    RC2_Transmit_PDO_Mapping_StatusWord_6041_00 : UINT;
    RC2_Transmit_PDO_Mapping_Position_actual_value_6064_00 : DINT;
    RC2_Transmit_PDO_Mapping_Mode_of_operation_display_6061_00 : SINT;
    RC2_Transmit_PDO_Mapping_Following_error_actual_valu_60F4_00 : DINT;
    RC2_Transmit_PDO_Mapping_Torque_actual_value_6077_00 : INT;
    RC2_Transmit_PDO_Mapping_Digital_inputs_60FD_00 : UDINT;
    RC2_Transmit_PDO_Mapping_Error_code_603F_00 : UINT;
    RC3_Receive_PDO_Mapping_ControlWord_6040_00 : UINT;
    RC3_Receive_PDO_Mapping_Target_Position_607A_00 : DINT;
    RC3_Receive_PDO_Mapping_Mode_of_operation_6060_00 : SINT;
    RC3_Receive_PDO_Mapping_Profile_velocity_6081_00 : UDINT;
    RC3_Receive_PDO_Mapping_Profile_acceleration_6083_00 : UDINT;
    RC3_Receive_PDO_Mapping_Profile_deceleration_6084_00 : UDINT;
    RC3_Receive_PDO_Mapping_Physical_outputs_60FE_01 : UDINT;
    RC3_Transmit_PDO_Mapping_StatusWord_6041_00 : UINT;
    RC3_Transmit_PDO_Mapping_Position_actual_value_6064_00 : DINT;
    RC3_Transmit_PDO_Mapping_Mode_of_operation_display_6061_00 : SINT;
    RC3_Transmit_PDO_Mapping_Following_error_actual_valu_60F4_00 : DINT;
    RC3_Transmit_PDO_Mapping_Torque_actual_value_6077_00 : INT;
    RC3_Transmit_PDO_Mapping_Digital_inputs_60FD_00 : UDINT;
    RC3_Transmit_PDO_Mapping_Error_code_603F_00 : UINT;
    RC4_Receive_PDO_Mapping_ControlWord_6040_00 : UINT;
    RC4_Receive_PDO_Mapping_Target_Position_607A_00 : DINT;
    RC4_Receive_PDO_Mapping_Mode_of_operation_6060_00 : SINT;
    RC4_Receive_PDO_Mapping_Profile_velocity_6081_00 : UDINT;
    RC4_Receive_PDO_Mapping_Profile_acceleration_6083_00 : UDINT;
    RC4_Receive_PDO_Mapping_Profile_deceleration_6084_00 : UDINT;
    RC4_Receive_PDO_Mapping_Physical_outputs_60FE_01 : UDINT;
    RC4_Transmit_PDO_Mapping_StatusWord_6041_00 : UINT;
    RC4_Transmit_PDO_Mapping_Position_actual_value_6064_00 : DINT;
    RC4_Transmit_PDO_Mapping_Mode_of_operation_display_6061_00 : SINT;
    RC4_Transmit_PDO_Mapping_Following_error_actual_valu_60F4_00 : DINT;
    RC4_Transmit_PDO_Mapping_Torque_actual_value_6077_00 : INT;
    RC4_Transmit_PDO_Mapping_Digital_inputs_60FD_00 : UDINT;
    RC4_Transmit_PDO_Mapping_Error_code_603F_00 : UINT;
    RC5_Receive_PDO_Mapping_ControlWord_6040_00 : UINT;
    RC5_Receive_PDO_Mapping_Target_Position_607A_00 : DINT;
    RC5_Receive_PDO_Mapping_Mode_of_operation_6060_00 : SINT;
    RC5_Receive_PDO_Mapping_Profile_velocity_6081_00 : UDINT;
    RC5_Receive_PDO_Mapping_Profile_acceleration_6083_00 : UDINT;
    RC5_Receive_PDO_Mapping_Profile_deceleration_6084_00 : UDINT;
    RC5_Receive_PDO_Mapping_Physical_outputs_60FE_01 : UDINT;
    RC5_Transmit_PDO_Mapping_StatusWord_6041_00 : UINT;
    RC5_Transmit_PDO_Mapping_Position_actual_value_6064_00 : DINT;
    RC5_Transmit_PDO_Mapping_Mode_of_operation_display_6061_00 : SINT;
    RC5_Transmit_PDO_Mapping_Following_error_actual_valu_60F4_00 : DINT;
    RC5_Transmit_PDO_Mapping_Torque_actual_value_6077_00 : INT;
    RC5_Transmit_PDO_Mapping_Digital_inputs_60FD_00 : UDINT;
    RC5_Transmit_PDO_Mapping_Error_code_603F_00 : UINT;
    RC6_Receive_PDO_Mapping_ControlWord_6040_00 : UINT;
    RC6_Receive_PDO_Mapping_ControlWord_6040_00_1 : UINT;
    RC6_Receive_PDO_Mapping_Target_Position_607A_00 : DINT;
    RC6_Receive_PDO_Mapping_Mode_of_operation_6060_00 : SINT;
    RC6_Receive_PDO_Mapping_Profile_velocity_6081_00 : UDINT;
    RC6_Receive_PDO_Mapping_Profile_acceleration_6083_00 : UDINT;
    RC6_Receive_PDO_Mapping_Profile_deceleration_6084_00 : UDINT;
    RC6_Receive_PDO_Mapping_Physical_outputs_60FE_01 : UDINT;
    RC6_Transmit_PDO_Mapping_StatusWord_6041_00 : UINT;
    RC6_Transmit_PDO_Mapping_Position_actual_value_6064_00 : DINT;
    RC6_Transmit_PDO_Mapping_Mode_of_operation_display_6061_00 : SINT;
    RC6_Transmit_PDO_Mapping_Following_error_actual_valu_60F4_00 : DINT;
    RC6_Transmit_PDO_Mapping_Torque_actual_value_6077_00 : INT;
    RC6_Transmit_PDO_Mapping_Digital_inputs_60FD_00 : UDINT;
    RC6_Transmit_PDO_Mapping_Error_code_603F_00 : UINT;
END_VAR
VAR_GLOBAL RETAIN
    RCON1_OUT : ARRAY[1..6] OF ST_RCON_Direct_OUT_Axis;  (* #RCON1 出力値; [2] #B(右側) NG1排出(上下); [3] #A(左側) SF/NG2仕分け(左右); [4] #B(右側) SF/NG2排出(送り); [5] #A(左側) SF/NG2排出(上下); [6] #B(右側) SF/NG2排出(上下); [1].Control.Pause 一時停止（安全停止とは別）（未接続）; [1] #A(左側) NG1排出(上下); [1].TargetPos_mm 目標位置 [mm]; [1].PositionBand_mm 位置決め幅 [mm]; [1].Speed_mm_s 指令速度 [mm/s]; [1].AccDec_G 加減速度 [G]; [1].PushLimit_pct 押付け制限 [%]（未使用）; [1].Control.Start 移動開始; [1].Control.Home 原点復帰（未接続）; [1].Control.Reset 異常リセット; [1].Control.ServoOn サーボON; [1].Control.InchingSelect インチング選択（OFF=ジョグ）; [1].Control.JogSpeedSelect ジョグ速度切替（未接続）; [1].Control.JogMinus 原点方向ジョグ（未接続）; [1].Control.JogPlus 反原点方向ジョグ（未接続）; [1].Control.GainSelect0 ゲイン選択0（未使用）; [1].Control.GainSelect1 ゲイン選択1（未使用）; [1].Control.PushEnable 押付け選択（OFF=位置決め）（未使用）; [1].Control.PushDirection 押付け方向（未使用）; [1].Control.RelativeMove 相対移動（OFF=絶対）（未使用）; [1].Control.BrakeRelease ブレーキ強制解除（落下注意）; [2].TargetPos_mm 目標位置 [mm]; [2].PositionBand_mm 位置決め幅 [mm]; [2].Speed_mm_s 指令速度 [mm/s]; [2].AccDec_G 加減速度 [G]; [2].PushLimit_pct 押付け制限 [%]（未使用）; [2].Control.Start 移動開始; [2].Control.Home 原点復帰（未接続）; [2].Control.Pause 一時停止（安全停止とは別）（未接続）; [2].Control.Reset 異常リセット; [2].Control.ServoOn サーボON; [2].Control.InchingSelect インチング選択（OFF=ジョグ）; [2].Control.JogSpeedSelect ジョグ速度切替（未接続）; [2].Control.JogMinus 原点方向ジョグ（未接続）; [2].Control.JogPlus 反原点方向ジョグ（未接続）; [2].Control.GainSelect0 ゲイン選択0（未使用）; [2].Control.GainSelect1 ゲイン選択1（未使用）; [2].Control.PushEnable 押付け選択（OFF=位置決め）（未使用）; [2].Control.PushDirection 押付け方向（未使用）; [2].Control.RelativeMove 相対移動（OFF=絶対）（未使用）; [2].Control.BrakeRelease ブレーキ強制解除（落下注意）; [3].TargetPos_mm 目標位置 [mm]; [3].PositionBand_mm 位置決め幅 [mm]; [3].Speed_mm_s 指令速度 [mm/s]; [3].AccDec_G 加減速度 [G]; [3].PushLimit_pct 押付け制限 [%]（未使用）; [3].Control.Start 移動開始; [3].Control.Home 原点復帰（未接続）; [3].Control.Pause 一時停止（安全停止とは別）（未接続）; [3].Control.Reset 異常リセット; [3].Control.ServoOn サーボON; [3].Control.InchingSelect インチング選択（OFF=ジョグ）; [3].Control.JogSpeedSelect ジョグ速度切替（未接続）; [3].Control.JogMinus 原点方向ジョグ（未接続）; [3].Control.JogPlus 反原点方向ジョグ（未接続）; [3].Control.GainSelect0 ゲイン選択0（未使用）; [3].Control.GainSelect1 ゲイン選択1（未使用）; [3].Control.PushEnable 押付け選択（OFF=位置決め）（未使用）; [3].Control.PushDirection 押付け方向（未使用）; [3].Control.RelativeMove 相対移動（OFF=絶対）（未使用）; [3].Control.BrakeRelease ブレーキ強制解除（落下注意）; [4].TargetPos_mm 目標位置 [mm]; [4].PositionBand_mm 位置決め幅 [mm]; [4].Speed_mm_s 指令速度 [mm/s]; [4].AccDec_G 加減速度 [G]; [4].PushLimit_pct 押付け制限 [%]（未使用）; [4].Control.Start 移動開始; [4].Control.Home 原点復帰（未接続）; [4].Control.Pause 一時停止（安全停止とは別）（未接続）; [4].Control.Reset 異常リセット; [4].Control.ServoOn サーボON; [4].Control.InchingSelect インチング選択（OFF=ジョグ）; [4].Control.JogSpeedSelect ジョグ速度切替（未接続）; [4].Control.JogMinus 原点方向ジョグ（未接続）; [4].Control.JogPlus 反原点方向ジョグ（未接続）; [4].Control.GainSelect0 ゲイン選択0（未使用）; [4].Control.GainSelect1 ゲイン選択1（未使用）; [4].Control.PushEnable 押付け選択（OFF=位置決め）（未使用）; [4].Control.PushDirection 押付け方向（未使用）; [4].Control.RelativeMove 相対移動（OFF=絶対）（未使用）; [4].Control.BrakeRelease ブレーキ強制解除（落下注意）; [5].TargetPos_mm 目標位置 [mm]; [5].PositionBand_mm 位置決め幅 [mm]; [5].Speed_mm_s 指令速度 [mm/s]; [5].AccDec_G 加減速度 [G]; [5].PushLimit_pct 押付け制限 [%]（未使用）; [5].Control.Start 移動開始; [5].Control.Home 原点復帰（未接続）; [5].Control.Pause 一時停止（安全停止とは別）（未接続）; [5].Control.Reset 異常リセット; [5].Control.ServoOn サーボON; [5].Control.InchingSelect インチング選択（OFF=ジョグ）; [5].Control.JogSpeedSelect ジョグ速度切替（未接続）; [5].Control.JogMinus 原点方向ジョグ（未接続）; [5].Control.JogPlus 反原点方向ジョグ（未接続）; [5].Control.GainSelect0 ゲイン選択0（未使用）; [5].Control.GainSelect1 ゲイン選択1（未使用）; [5].Control.PushEnable 押付け選択（OFF=位置決め）（未使用）; [5].Control.PushDirection 押付け方向（未使用）; [5].Control.RelativeMove 相対移動（OFF=絶対）（未使用）; [5].Control.BrakeRelease ブレーキ強制解除（落下注意）; [6].TargetPos_mm 目標位置 [mm]; [6].PositionBand_mm 位置決め幅 [mm]; [6].Speed_mm_s 指令速度 [mm/s]; [6].AccDec_G 加減速度 [G]; [6].PushLimit_pct 押付け制限 [%]（未使用）; [6].Control.Start 移動開始; [6].Control.Home 原点復帰（未接続）; [6].Control.Pause 一時停止（安全停止とは別）（未接続）; [6].Control.Reset 異常リセット; [6].Control.ServoOn サーボON; [6].Control.InchingSelect インチング選択（OFF=ジョグ）; [6].Control.JogSpeedSelect ジョグ速度切替（未接続）; [6].Control.JogMinus 原点方向ジョグ（未接続）; [6].Control.JogPlus 反原点方向ジョグ（未接続）; [6].Control.GainSelect0 ゲイン選択0（未使用）; [6].Control.GainSelect1 ゲイン選択1（未使用）; [6].Control.PushEnable 押付け選択（OFF=位置決め）（未使用）; [6].Control.PushDirection 押付け方向（未使用）; [6].Control.RelativeMove 相対移動（OFF=絶対）（未使用）; [6].Control.BrakeRelease ブレーキ強制解除（落下注意） *)
    RCON1_IN : ARRAY[1..6] OF ST_RCON_Direct_IN_Axis;  (* #RCON1 入力値; [1] #A(左側) NG1排出(上下); [2] #B(右側) NG1排出(上下); [3] #A(左側) SF/NG2仕分け(左右); [4] #B(右側) SF/NG2排出(送り); [5] #A(左側) SF/NG2排出(上下); [6] #B(右側) SF/NG2排出(上下); [1].ActualPos_mm 現在位置 [mm]; [1].Current_mA 指令電流 [mA]; [1].ActualSpeed_mm_s 現在速度 [mm/s]; [1].AlarmCode 異常コード; [1].DataValid 入力有効（安全許可とは別）; [1].Status.PositionDone 位置決め完了; [1].Status.HomeDone 原点復帰完了; [1].Status.Moving 移動中; [1].Status.Alarm 軸異常; [1].Status.ServoReady サーボON状態; [1].Status.PushMiss 押付け空振り（未使用）; [1].Status.OverloadWarning 過負荷警告; [1].Status.CommandDone 指令完了（空振り含む）; [1].Status.Zone1 ゾーン1内; [1].Status.Zone2 ゾーン2内; [1].Status.ControllerReady 準備完了; [1].Status.EmergencyStop 非常停止状態（監視）; [2].ActualPos_mm 現在位置 [mm]; [2].Current_mA 指令電流 [mA]; [2].ActualSpeed_mm_s 現在速度 [mm/s]; [2].AlarmCode 異常コード; [2].DataValid 入力有効（安全許可とは別）; [2].Status.PositionDone 位置決め完了; [2].Status.HomeDone 原点復帰完了; [2].Status.Moving 移動中; [2].Status.Alarm 軸異常; [2].Status.ServoReady サーボON状態; [2].Status.PushMiss 押付け空振り（未使用）; [2].Status.OverloadWarning 過負荷警告; [2].Status.CommandDone 指令完了（空振り含む）; [2].Status.Zone1 ゾーン1内; [2].Status.Zone2 ゾーン2内; [2].Status.ControllerReady 準備完了; [2].Status.EmergencyStop 非常停止状態（監視）; [3].ActualPos_mm 現在位置 [mm]; [3].Current_mA 指令電流 [mA]; [3].ActualSpeed_mm_s 現在速度 [mm/s]; [3].AlarmCode 異常コード; [3].DataValid 入力有効（安全許可とは別）; [3].Status.PositionDone 位置決め完了; [3].Status.HomeDone 原点復帰完了; [3].Status.Moving 移動中; [3].Status.Alarm 軸異常; [3].Status.ServoReady サーボON状態; [3].Status.PushMiss 押付け空振り（未使用）; [3].Status.OverloadWarning 過負荷警告; [3].Status.CommandDone 指令完了（空振り含む）; [3].Status.Zone1 ゾーン1内; [3].Status.Zone2 ゾーン2内; [3].Status.ControllerReady 準備完了; [3].Status.EmergencyStop 非常停止状態（監視）; [4].ActualPos_mm 現在位置 [mm]; [4].Current_mA 指令電流 [mA]; [4].ActualSpeed_mm_s 現在速度 [mm/s]; [4].AlarmCode 異常コード; [4].DataValid 入力有効（安全許可とは別）; [4].Status.PositionDone 位置決め完了; [4].Status.HomeDone 原点復帰完了; [4].Status.Moving 移動中; [4].Status.Alarm 軸異常; [4].Status.ServoReady サーボON状態; [4].Status.PushMiss 押付け空振り（未使用）; [4].Status.OverloadWarning 過負荷警告; [4].Status.CommandDone 指令完了（空振り含む）; [4].Status.Zone1 ゾーン1内; [4].Status.Zone2 ゾーン2内; [4].Status.ControllerReady 準備完了; [4].Status.EmergencyStop 非常停止状態（監視）; [5].ActualPos_mm 現在位置 [mm]; [5].Current_mA 指令電流 [mA]; [5].ActualSpeed_mm_s 現在速度 [mm/s]; [5].AlarmCode 異常コード; [5].DataValid 入力有効（安全許可とは別）; [5].Status.PositionDone 位置決め完了; [5].Status.HomeDone 原点復帰完了; [5].Status.Moving 移動中; [5].Status.Alarm 軸異常; [5].Status.ServoReady サーボON状態; [5].Status.PushMiss 押付け空振り（未使用）; [5].Status.OverloadWarning 過負荷警告; [5].Status.CommandDone 指令完了（空振り含む）; [5].Status.Zone1 ゾーン1内; [5].Status.Zone2 ゾーン2内; [5].Status.ControllerReady 準備完了; [5].Status.EmergencyStop 非常停止状態（監視）; [6].ActualPos_mm 現在位置 [mm]; [6].Current_mA 指令電流 [mA]; [6].ActualSpeed_mm_s 現在速度 [mm/s]; [6].AlarmCode 異常コード; [6].DataValid 入力有効（安全許可とは別）; [6].Status.PositionDone 位置決め完了; [6].Status.HomeDone 原点復帰完了; [6].Status.Moving 移動中; [6].Status.Alarm 軸異常; [6].Status.ServoReady サーボON状態; [6].Status.PushMiss 押付け空振り（未使用）; [6].Status.OverloadWarning 過負荷警告; [6].Status.CommandDone 指令完了（空振り含む）; [6].Status.Zone1 ゾーン1内; [6].Status.Zone2 ゾーン2内; [6].Status.ControllerReady 準備完了; [6].Status.EmergencyStop 非常停止状態（監視） *)
END_VAR
VAR_GLOBAL
    RCON1_SpeedUnit_mm_s : LREAL;  (* 速度単位 [mm/s/カウント]（1.0/0.1） *)
    RCON1_OUT_GwControl0Raw : UINT;  (* 未割付・不使用 OUT00 共通制御（MON/RTE） *)
    RCON1_OUT_GwControl1ReservedRaw : UINT;  (* 未割付・不使用 OUT01 予約（書込禁止） *)
    RCON1_OUT_ReservedOut02Raw : UINT;  (* 未割付・不使用 OUT02 予約（書込禁止） *)
    RCON1_OUT_ReservedOut03Raw : UINT;  (* 未割付・不使用 OUT03 予約（書込禁止） *)
    RCON1_OUT_ReservedOut04Raw : UINT;  (* 未割付・不使用 OUT04 予約（書込禁止） *)
    RCON1_OUT_ReservedOut05Raw : UINT;  (* 未割付・不使用 OUT05 予約（書込禁止） *)
    RCON1_OUT_ReservedOut06Raw : UINT;  (* 未割付・不使用 OUT06 予約（書込禁止） *)
    RCON1_OUT_ReservedOut07Raw : UINT;  (* 未割付・不使用 OUT07 予約（書込禁止） *)
    RCON1_OUT_Axis1_TargetPosLoRaw : UINT;  (* 未割付・不使用 OUT08 1軸目 目標位置 下位 [0.01mm] *)
    RCON1_OUT_Axis1_TargetPosHiRaw : UINT;  (* 未割付・不使用 OUT09 1軸目 目標位置 上位 [0.01mm] *)
    RCON1_OUT_Axis1_PositionBandLoRaw : UINT;  (* 未割付・不使用 OUT10 1軸目 位置決め幅 下位 [0.01mm] *)
    RCON1_OUT_Axis1_PositionBandHiRaw : UINT;  (* 未割付・不使用 OUT11 1軸目 位置決め幅 上位 [0.01mm] *)
    RCON1_OUT_Axis1_SpeedRaw : UINT;  (* 未割付・不使用 OUT12 1軸目 速度指令 [実機単位] *)
    RCON1_OUT_Axis1_AccDecRaw : UINT;  (* 未割付・不使用 OUT13 1軸目 共通加減速 [0.01G] *)
    RCON1_OUT_Axis1_PushLimitRaw : UINT;  (* 未割付・不使用 OUT14 1軸目 押付け制限 [255=100%] *)
    RCON1_OUT_Axis1_ControlRaw : UINT;  (* 未割付・不使用 OUT15 1軸目 制御信号（DSTR/SON等） *)
    RCON1_OUT_Axis2_TargetPosLoRaw : UINT;  (* 未割付・不使用 OUT16 2軸目 目標位置 下位 [0.01mm] *)
    RCON1_OUT_Axis2_TargetPosHiRaw : UINT;  (* 未割付・不使用 OUT17 2軸目 目標位置 上位 [0.01mm] *)
    RCON1_OUT_Axis2_PositionBandLoRaw : UINT;  (* 未割付・不使用 OUT18 2軸目 位置決め幅 下位 [0.01mm] *)
    RCON1_OUT_Axis2_PositionBandHiRaw : UINT;  (* 未割付・不使用 OUT19 2軸目 位置決め幅 上位 [0.01mm] *)
    RCON1_OUT_Axis2_SpeedRaw : UINT;  (* 未割付・不使用 OUT20 2軸目 速度指令 [実機単位] *)
    RCON1_OUT_Axis2_AccDecRaw : UINT;  (* 未割付・不使用 OUT21 2軸目 共通加減速 [0.01G] *)
    RCON1_OUT_Axis2_PushLimitRaw : UINT;  (* 未割付・不使用 OUT22 2軸目 押付け制限 [255=100%] *)
    RCON1_OUT_Axis2_ControlRaw : UINT;  (* 未割付・不使用 OUT23 2軸目 制御信号（DSTR/SON等） *)
    RCON1_OUT_Axis3_TargetPosLoRaw : UINT;  (* 未割付・不使用 OUT24 3軸目 目標位置 下位 [0.01mm] *)
    RCON1_OUT_Axis3_TargetPosHiRaw : UINT;  (* 未割付・不使用 OUT25 3軸目 目標位置 上位 [0.01mm] *)
    RCON1_OUT_Axis3_PositionBandLoRaw : UINT;  (* 未割付・不使用 OUT26 3軸目 位置決め幅 下位 [0.01mm] *)
    RCON1_OUT_Axis3_PositionBandHiRaw : UINT;  (* 未割付・不使用 OUT27 3軸目 位置決め幅 上位 [0.01mm] *)
    RCON1_OUT_Axis3_SpeedRaw : UINT;  (* 未割付・不使用 OUT28 3軸目 速度指令 [実機単位] *)
    RCON1_OUT_Axis3_AccDecRaw : UINT;  (* 未割付・不使用 OUT29 3軸目 共通加減速 [0.01G] *)
    RCON1_OUT_Axis3_PushLimitRaw : UINT;  (* 未割付・不使用 OUT30 3軸目 押付け制限 [255=100%] *)
    RCON1_OUT_Axis3_ControlRaw : UINT;  (* 未割付・不使用 OUT31 3軸目 制御信号（DSTR/SON等） *)
    RCON1_OUT_Axis4_TargetPosLoRaw : UINT;  (* 未割付・不使用 OUT32 4軸目 目標位置 下位 [0.01mm] *)
    RCON1_OUT_Axis4_TargetPosHiRaw : UINT;  (* 未割付・不使用 OUT33 4軸目 目標位置 上位 [0.01mm] *)
    RCON1_OUT_Axis4_PositionBandLoRaw : UINT;  (* 未割付・不使用 OUT34 4軸目 位置決め幅 下位 [0.01mm] *)
    RCON1_OUT_Axis4_PositionBandHiRaw : UINT;  (* 未割付・不使用 OUT35 4軸目 位置決め幅 上位 [0.01mm] *)
    RCON1_OUT_Axis4_SpeedRaw : UINT;  (* 未割付・不使用 OUT36 4軸目 速度指令 [実機単位] *)
    RCON1_OUT_Axis4_AccDecRaw : UINT;  (* 未割付・不使用 OUT37 4軸目 共通加減速 [0.01G] *)
    RCON1_OUT_Axis4_PushLimitRaw : UINT;  (* 未割付・不使用 OUT38 4軸目 押付け制限 [255=100%] *)
    RCON1_OUT_Axis4_ControlRaw : UINT;  (* 未割付・不使用 OUT39 4軸目 制御信号（DSTR/SON等） *)
    RCON1_OUT_Axis5_TargetPosLoRaw : UINT;  (* 未割付・不使用 OUT40 5軸目 目標位置 下位 [0.01mm] *)
    RCON1_OUT_Axis5_TargetPosHiRaw : UINT;  (* 未割付・不使用 OUT41 5軸目 目標位置 上位 [0.01mm] *)
    RCON1_OUT_Axis5_PositionBandLoRaw : UINT;  (* 未割付・不使用 OUT42 5軸目 位置決め幅 下位 [0.01mm] *)
    RCON1_OUT_Axis5_PositionBandHiRaw : UINT;  (* 未割付・不使用 OUT43 5軸目 位置決め幅 上位 [0.01mm] *)
    RCON1_OUT_Axis5_SpeedRaw : UINT;  (* 未割付・不使用 OUT44 5軸目 速度指令 [実機単位] *)
    RCON1_OUT_Axis5_AccDecRaw : UINT;  (* 未割付・不使用 OUT45 5軸目 共通加減速 [0.01G] *)
    RCON1_OUT_Axis5_PushLimitRaw : UINT;  (* 未割付・不使用 OUT46 5軸目 押付け制限 [255=100%] *)
    RCON1_OUT_Axis5_ControlRaw : UINT;  (* 未割付・不使用 OUT47 5軸目 制御信号（DSTR/SON等） *)
    RCON1_OUT_Axis6_TargetPosLoRaw : UINT;  (* 未割付・不使用 OUT48 6軸目 目標位置 下位 [0.01mm] *)
    RCON1_OUT_Axis6_TargetPosHiRaw : UINT;  (* 未割付・不使用 OUT49 6軸目 目標位置 上位 [0.01mm] *)
    RCON1_OUT_Axis6_PositionBandLoRaw : UINT;  (* 未割付・不使用 OUT50 6軸目 位置決め幅 下位 [0.01mm] *)
    RCON1_OUT_Axis6_PositionBandHiRaw : UINT;  (* 未割付・不使用 OUT51 6軸目 位置決め幅 上位 [0.01mm] *)
    RCON1_OUT_Axis6_SpeedRaw : UINT;  (* 未割付・不使用 OUT52 6軸目 速度指令 [実機単位] *)
    RCON1_OUT_Axis6_AccDecRaw : UINT;  (* 未割付・不使用 OUT53 6軸目 共通加減速 [0.01G] *)
    RCON1_OUT_Axis6_PushLimitRaw : UINT;  (* 未割付・不使用 OUT54 6軸目 押付け制限 [255=100%] *)
    RCON1_OUT_Axis6_ControlRaw : UINT;  (* 未割付・不使用 OUT55 6軸目 制御信号（DSTR/SON等） *)
    RCON1_IN_GwStatus0Raw : UINT;  (* 未割付・不使用 IN00 GW状態 *)
    RCON1_IN_AxisLinkStatusRaw : UINT;  (* 未割付・不使用 IN01 軸リンク状態 *)
    RCON1_IN_PowerStatus0Raw : UINT;  (* 未割付・不使用 IN02 電源状態0 *)
    RCON1_IN_PowerStatus1Raw : UINT;  (* 未割付・不使用 IN03 電源状態1 *)
    RCON1_IN_PowerStatus2Raw : UINT;  (* 未割付・不使用 IN04 電源状態2 *)
    RCON1_IN_PowerStatus3Raw : UINT;  (* 未割付・不使用 IN05 電源状態3 *)
    RCON1_IN_PowerStatus4MaintenanceRaw : UINT;  (* 未割付・不使用 IN06 電源状態4（構成依存） *)
    RCON1_IN_ReservedIn07Raw : UINT;  (* 未割付・不使用 IN07 予約（使用禁止） *)
    RCON1_IN_Axis1_ActualPosLoRaw : UINT;  (* 未割付・不使用 IN08 1軸目 現在位置 下位 [0.01mm] *)
    RCON1_IN_Axis1_ActualPosHiRaw : UINT;  (* 未割付・不使用 IN09 1軸目 現在位置 上位 [0.01mm] *)
    RCON1_IN_Axis1_CurrentLoRaw : UINT;  (* 未割付・不使用 IN10 1軸目 指令電流 下位 [mA] *)
    RCON1_IN_Axis1_CurrentHiRaw : UINT;  (* 未割付・不使用 IN11 1軸目 指令電流 上位 [mA] *)
    RCON1_IN_Axis1_ActualSpeedRaw : UINT;  (* 未割付・不使用 IN12 1軸目 現在速度 [実機単位・符号付き] *)
    RCON1_IN_Axis1_ReservedInRaw : UINT;  (* 未割付・不使用 IN13 1軸目 予約（使用禁止） *)
    RCON1_IN_Axis1_AlarmCodeRaw : UINT;  (* 未割付・不使用 IN14 1軸目 軸異常コード *)
    RCON1_IN_Axis1_StatusRaw : UINT;  (* 未割付・不使用 IN15 1軸目 状態信号（PEND/SV等） *)
    RCON1_IN_Axis2_ActualPosLoRaw : UINT;  (* 未割付・不使用 IN16 2軸目 現在位置 下位 [0.01mm] *)
    RCON1_IN_Axis2_ActualPosHiRaw : UINT;  (* 未割付・不使用 IN17 2軸目 現在位置 上位 [0.01mm] *)
    RCON1_IN_Axis2_CurrentLoRaw : UINT;  (* 未割付・不使用 IN18 2軸目 指令電流 下位 [mA] *)
    RCON1_IN_Axis2_CurrentHiRaw : UINT;  (* 未割付・不使用 IN19 2軸目 指令電流 上位 [mA] *)
    RCON1_IN_Axis2_ActualSpeedRaw : UINT;  (* 未割付・不使用 IN20 2軸目 現在速度 [実機単位・符号付き] *)
    RCON1_IN_Axis2_ReservedInRaw : UINT;  (* 未割付・不使用 IN21 2軸目 予約（使用禁止） *)
    RCON1_IN_Axis2_AlarmCodeRaw : UINT;  (* 未割付・不使用 IN22 2軸目 軸異常コード *)
    RCON1_IN_Axis2_StatusRaw : UINT;  (* 未割付・不使用 IN23 2軸目 状態信号（PEND/SV等） *)
    RCON1_IN_Axis3_ActualPosLoRaw : UINT;  (* 未割付・不使用 IN24 3軸目 現在位置 下位 [0.01mm] *)
    RCON1_IN_Axis3_ActualPosHiRaw : UINT;  (* 未割付・不使用 IN25 3軸目 現在位置 上位 [0.01mm] *)
    RCON1_IN_Axis3_CurrentLoRaw : UINT;  (* 未割付・不使用 IN26 3軸目 指令電流 下位 [mA] *)
    RCON1_IN_Axis3_CurrentHiRaw : UINT;  (* 未割付・不使用 IN27 3軸目 指令電流 上位 [mA] *)
    RCON1_IN_Axis3_ActualSpeedRaw : UINT;  (* 未割付・不使用 IN28 3軸目 現在速度 [実機単位・符号付き] *)
    RCON1_IN_Axis3_ReservedInRaw : UINT;  (* 未割付・不使用 IN29 3軸目 予約（使用禁止） *)
    RCON1_IN_Axis3_AlarmCodeRaw : UINT;  (* 未割付・不使用 IN30 3軸目 軸異常コード *)
    RCON1_IN_Axis3_StatusRaw : UINT;  (* 未割付・不使用 IN31 3軸目 状態信号（PEND/SV等） *)
    RCON1_IN_Axis4_ActualPosLoRaw : UINT;  (* 未割付・不使用 IN32 4軸目 現在位置 下位 [0.01mm] *)
    RCON1_IN_Axis4_ActualPosHiRaw : UINT;  (* 未割付・不使用 IN33 4軸目 現在位置 上位 [0.01mm] *)
    RCON1_IN_Axis4_CurrentLoRaw : UINT;  (* 未割付・不使用 IN34 4軸目 指令電流 下位 [mA] *)
    RCON1_IN_Axis4_CurrentHiRaw : UINT;  (* 未割付・不使用 IN35 4軸目 指令電流 上位 [mA] *)
    RCON1_IN_Axis4_ActualSpeedRaw : UINT;  (* 未割付・不使用 IN36 4軸目 現在速度 [実機単位・符号付き] *)
    RCON1_IN_Axis4_ReservedInRaw : UINT;  (* 未割付・不使用 IN37 4軸目 予約（使用禁止） *)
    RCON1_IN_Axis4_AlarmCodeRaw : UINT;  (* 未割付・不使用 IN38 4軸目 軸異常コード *)
    RCON1_IN_Axis4_StatusRaw : UINT;  (* 未割付・不使用 IN39 4軸目 状態信号（PEND/SV等） *)
    RCON1_IN_Axis5_ActualPosLoRaw : UINT;  (* 未割付・不使用 IN40 5軸目 現在位置 下位 [0.01mm] *)
    RCON1_IN_Axis5_ActualPosHiRaw : UINT;  (* 未割付・不使用 IN41 5軸目 現在位置 上位 [0.01mm] *)
    RCON1_IN_Axis5_CurrentLoRaw : UINT;  (* 未割付・不使用 IN42 5軸目 指令電流 下位 [mA] *)
    RCON1_IN_Axis5_CurrentHiRaw : UINT;  (* 未割付・不使用 IN43 5軸目 指令電流 上位 [mA] *)
    RCON1_IN_Axis5_ActualSpeedRaw : UINT;  (* 未割付・不使用 IN44 5軸目 現在速度 [実機単位・符号付き] *)
    RCON1_IN_Axis5_ReservedInRaw : UINT;  (* 未割付・不使用 IN45 5軸目 予約（使用禁止） *)
    RCON1_IN_Axis5_AlarmCodeRaw : UINT;  (* 未割付・不使用 IN46 5軸目 軸異常コード *)
    RCON1_IN_Axis5_StatusRaw : UINT;  (* 未割付・不使用 IN47 5軸目 状態信号（PEND/SV等） *)
    RCON1_IN_Axis6_ActualPosLoRaw : UINT;  (* 未割付・不使用 IN48 6軸目 現在位置 下位 [0.01mm] *)
    RCON1_IN_Axis6_ActualPosHiRaw : UINT;  (* 未割付・不使用 IN49 6軸目 現在位置 上位 [0.01mm] *)
    RCON1_IN_Axis6_CurrentLoRaw : UINT;  (* 未割付・不使用 IN50 6軸目 指令電流 下位 [mA] *)
    RCON1_IN_Axis6_CurrentHiRaw : UINT;  (* 未割付・不使用 IN51 6軸目 指令電流 上位 [mA] *)
    RCON1_IN_Axis6_ActualSpeedRaw : UINT;  (* 未割付・不使用 IN52 6軸目 現在速度 [実機単位・符号付き] *)
    RCON1_IN_Axis6_ReservedInRaw : UINT;  (* 未割付・不使用 IN53 6軸目 予約（使用禁止） *)
    RCON1_IN_Axis6_AlarmCodeRaw : UINT;  (* 未割付・不使用 IN54 6軸目 軸異常コード *)
END_VAR
VAR_GLOBAL RETAIN
    RCON1_IN_Axis6_StatusRaw : UINT;  (* 未割付・不使用 IN55 6軸目 状態信号（PEND/SV等） *)
    RCON2_OUT : ARRAY[1..5] OF ST_RCON_Direct_OUT_Axis;  (* #RCON2 出力値; [1] 1軸目（No.0）出力指令; [2] 2軸目（No.1）出力指令; [3] 3軸目（No.2）出力指令; [4] 4軸目（No.3）出力指令; [5] 5軸目（No.4）出力指令 *)
END_VAR
VAR_GLOBAL
    RCON2_IN : ARRAY[1..5] OF ST_RCON_Direct_IN_Axis;  (* #RCON2 入力値; [1] 1軸目（No.0）入力情報; [2] 2軸目（No.1）入力情報; [3] 3軸目（No.2）入力情報; [4] 4軸目（No.3）入力情報; [5] 5軸目（No.4）入力情報 *)
    RCON2_SpeedUnit_mm_s : LREAL;  (* 速度単位 [mm/s/カウント]（1.0/0.1） *)
    RCON2_OUT_GwControl0Raw : UINT;  (* 未割付・不使用 OUT00 共通制御（MON/RTE） *)
    RCON2_OUT_GwControl1ReservedRaw : UINT;  (* 未割付・不使用 OUT01 予約（書込禁止） *)
    RCON2_OUT_ReservedOut02Raw : UINT;  (* 未割付・不使用 OUT02 予約（書込禁止） *)
    RCON2_OUT_ReservedOut03Raw : UINT;  (* 未割付・不使用 OUT03 予約（書込禁止） *)
    RCON2_OUT_ReservedOut04Raw : UINT;  (* 未割付・不使用 OUT04 予約（書込禁止） *)
    RCON2_OUT_ReservedOut05Raw : UINT;  (* 未割付・不使用 OUT05 予約（書込禁止） *)
    RCON2_OUT_ReservedOut06Raw : UINT;  (* 未割付・不使用 OUT06 予約（書込禁止） *)
    RCON2_OUT_ReservedOut07Raw : UINT;  (* 未割付・不使用 OUT07 予約（書込禁止） *)
    RCON2_OUT_Axis1_TargetPosLoRaw : UINT;  (* 未割付・不使用 OUT08 1軸目 目標位置 下位 [0.01mm] *)
    RCON2_OUT_Axis1_TargetPosHiRaw : UINT;  (* 未割付・不使用 OUT09 1軸目 目標位置 上位 [0.01mm] *)
    RCON2_OUT_Axis1_PositionBandLoRaw : UINT;  (* 未割付・不使用 OUT10 1軸目 位置決め幅 下位 [0.01mm] *)
    RCON2_OUT_Axis1_PositionBandHiRaw : UINT;  (* 未割付・不使用 OUT11 1軸目 位置決め幅 上位 [0.01mm] *)
    RCON2_OUT_Axis1_SpeedRaw : UINT;  (* 未割付・不使用 OUT12 1軸目 速度指令 [実機単位] *)
    RCON2_OUT_Axis1_AccDecRaw : UINT;  (* 未割付・不使用 OUT13 1軸目 共通加減速 [0.01G] *)
    RCON2_OUT_Axis1_PushLimitRaw : UINT;  (* 未割付・不使用 OUT14 1軸目 押付け制限 [255=100%] *)
    RCON2_OUT_Axis1_ControlRaw : UINT;  (* 未割付・不使用 OUT15 1軸目 制御信号（DSTR/SON等） *)
    RCON2_OUT_Axis2_TargetPosLoRaw : UINT;  (* 未割付・不使用 OUT16 2軸目 目標位置 下位 [0.01mm] *)
    RCON2_OUT_Axis2_TargetPosHiRaw : UINT;  (* 未割付・不使用 OUT17 2軸目 目標位置 上位 [0.01mm] *)
    RCON2_OUT_Axis2_PositionBandLoRaw : UINT;  (* 未割付・不使用 OUT18 2軸目 位置決め幅 下位 [0.01mm] *)
    RCON2_OUT_Axis2_PositionBandHiRaw : UINT;  (* 未割付・不使用 OUT19 2軸目 位置決め幅 上位 [0.01mm] *)
    RCON2_OUT_Axis2_SpeedRaw : UINT;  (* 未割付・不使用 OUT20 2軸目 速度指令 [実機単位] *)
    RCON2_OUT_Axis2_AccDecRaw : UINT;  (* 未割付・不使用 OUT21 2軸目 共通加減速 [0.01G] *)
    RCON2_OUT_Axis2_PushLimitRaw : UINT;  (* 未割付・不使用 OUT22 2軸目 押付け制限 [255=100%] *)
    RCON2_OUT_Axis2_ControlRaw : UINT;  (* 未割付・不使用 OUT23 2軸目 制御信号（DSTR/SON等） *)
    RCON2_OUT_Axis3_TargetPosLoRaw : UINT;  (* 未割付・不使用 OUT24 3軸目 目標位置 下位 [0.01mm] *)
    RCON2_OUT_Axis3_TargetPosHiRaw : UINT;  (* 未割付・不使用 OUT25 3軸目 目標位置 上位 [0.01mm] *)
    RCON2_OUT_Axis3_PositionBandLoRaw : UINT;  (* 未割付・不使用 OUT26 3軸目 位置決め幅 下位 [0.01mm] *)
    RCON2_OUT_Axis3_PositionBandHiRaw : UINT;  (* 未割付・不使用 OUT27 3軸目 位置決め幅 上位 [0.01mm] *)
    RCON2_OUT_Axis3_SpeedRaw : UINT;  (* 未割付・不使用 OUT28 3軸目 速度指令 [実機単位] *)
    RCON2_OUT_Axis3_AccDecRaw : UINT;  (* 未割付・不使用 OUT29 3軸目 共通加減速 [0.01G] *)
    RCON2_OUT_Axis3_PushLimitRaw : UINT;  (* 未割付・不使用 OUT30 3軸目 押付け制限 [255=100%] *)
    RCON2_OUT_Axis3_ControlRaw : UINT;  (* 未割付・不使用 OUT31 3軸目 制御信号（DSTR/SON等） *)
    RCON2_OUT_Axis4_TargetPosLoRaw : UINT;  (* 未割付・不使用 OUT32 4軸目 目標位置 下位 [0.01mm] *)
    RCON2_OUT_Axis4_TargetPosHiRaw : UINT;  (* 未割付・不使用 OUT33 4軸目 目標位置 上位 [0.01mm] *)
    RCON2_OUT_Axis4_PositionBandLoRaw : UINT;  (* 未割付・不使用 OUT34 4軸目 位置決め幅 下位 [0.01mm] *)
    RCON2_OUT_Axis4_PositionBandHiRaw : UINT;  (* 未割付・不使用 OUT35 4軸目 位置決め幅 上位 [0.01mm] *)
    RCON2_OUT_Axis4_SpeedRaw : UINT;  (* 未割付・不使用 OUT36 4軸目 速度指令 [実機単位] *)
    RCON2_OUT_Axis4_AccDecRaw : UINT;  (* 未割付・不使用 OUT37 4軸目 共通加減速 [0.01G] *)
    RCON2_OUT_Axis4_PushLimitRaw : UINT;  (* 未割付・不使用 OUT38 4軸目 押付け制限 [255=100%] *)
    RCON2_OUT_Axis4_ControlRaw : UINT;  (* 未割付・不使用 OUT39 4軸目 制御信号（DSTR/SON等） *)
    RCON2_OUT_Axis5_TargetPosLoRaw : UINT;  (* 未割付・不使用 OUT40 5軸目 目標位置 下位 [0.01mm] *)
    RCON2_OUT_Axis5_TargetPosHiRaw : UINT;  (* 未割付・不使用 OUT41 5軸目 目標位置 上位 [0.01mm] *)
    RCON2_OUT_Axis5_PositionBandLoRaw : UINT;  (* 未割付・不使用 OUT42 5軸目 位置決め幅 下位 [0.01mm] *)
    RCON2_OUT_Axis5_PositionBandHiRaw : UINT;  (* 未割付・不使用 OUT43 5軸目 位置決め幅 上位 [0.01mm] *)
    RCON2_OUT_Axis5_SpeedRaw : UINT;  (* 未割付・不使用 OUT44 5軸目 速度指令 [実機単位] *)
    RCON2_OUT_Axis5_AccDecRaw : UINT;  (* 未割付・不使用 OUT45 5軸目 共通加減速 [0.01G] *)
    RCON2_OUT_Axis5_PushLimitRaw : UINT;  (* 未割付・不使用 OUT46 5軸目 押付け制限 [255=100%] *)
    RCON2_OUT_Axis5_ControlRaw : UINT;  (* 未割付・不使用 OUT47 5軸目 制御信号（DSTR/SON等） *)
    RCON2_IN_GwStatus0Raw : UINT;  (* 未割付・不使用 IN00 GW状態 *)
    RCON2_IN_AxisLinkStatusRaw : UINT;  (* 未割付・不使用 IN01 軸リンク状態 *)
    RCON2_IN_PowerStatus0Raw : UINT;  (* 未割付・不使用 IN02 電源状態0 *)
    RCON2_IN_PowerStatus1Raw : UINT;  (* 未割付・不使用 IN03 電源状態1 *)
    RCON2_IN_PowerStatus2Raw : UINT;  (* 未割付・不使用 IN04 電源状態2 *)
    RCON2_IN_PowerStatus3Raw : UINT;  (* 未割付・不使用 IN05 電源状態3 *)
    RCON2_IN_PowerStatus4MaintenanceRaw : UINT;  (* 未割付・不使用 IN06 電源状態4（構成依存） *)
    RCON2_IN_ReservedIn07Raw : UINT;  (* 未割付・不使用 IN07 予約（使用禁止） *)
    RCON2_IN_Axis1_ActualPosLoRaw : UINT;  (* 未割付・不使用 IN08 1軸目 現在位置 下位 [0.01mm] *)
    RCON2_IN_Axis1_ActualPosHiRaw : UINT;  (* 未割付・不使用 IN09 1軸目 現在位置 上位 [0.01mm] *)
    RCON2_IN_Axis1_CurrentLoRaw : UINT;  (* 未割付・不使用 IN10 1軸目 指令電流 下位 [mA] *)
    RCON2_IN_Axis1_CurrentHiRaw : UINT;  (* 未割付・不使用 IN11 1軸目 指令電流 上位 [mA] *)
    RCON2_IN_Axis1_ActualSpeedRaw : UINT;  (* 未割付・不使用 IN12 1軸目 現在速度 [実機単位・符号付き] *)
    RCON2_IN_Axis1_ReservedInRaw : UINT;  (* 未割付・不使用 IN13 1軸目 予約（使用禁止） *)
    RCON2_IN_Axis1_AlarmCodeRaw : UINT;  (* 未割付・不使用 IN14 1軸目 軸異常コード *)
    RCON2_IN_Axis1_StatusRaw : UINT;  (* 未割付・不使用 IN15 1軸目 状態信号（PEND/SV等） *)
    RCON2_IN_Axis2_ActualPosLoRaw : UINT;  (* 未割付・不使用 IN16 2軸目 現在位置 下位 [0.01mm] *)
    RCON2_IN_Axis2_ActualPosHiRaw : UINT;  (* 未割付・不使用 IN17 2軸目 現在位置 上位 [0.01mm] *)
    RCON2_IN_Axis2_CurrentLoRaw : UINT;  (* 未割付・不使用 IN18 2軸目 指令電流 下位 [mA] *)
    RCON2_IN_Axis2_CurrentHiRaw : UINT;  (* 未割付・不使用 IN19 2軸目 指令電流 上位 [mA] *)
    RCON2_IN_Axis2_ActualSpeedRaw : UINT;  (* 未割付・不使用 IN20 2軸目 現在速度 [実機単位・符号付き] *)
    RCON2_IN_Axis2_ReservedInRaw : UINT;  (* 未割付・不使用 IN21 2軸目 予約（使用禁止） *)
    RCON2_IN_Axis2_AlarmCodeRaw : UINT;  (* 未割付・不使用 IN22 2軸目 軸異常コード *)
    RCON2_IN_Axis2_StatusRaw : UINT;  (* 未割付・不使用 IN23 2軸目 状態信号（PEND/SV等） *)
    RCON2_IN_Axis3_ActualPosLoRaw : UINT;  (* 未割付・不使用 IN24 3軸目 現在位置 下位 [0.01mm] *)
    RCON2_IN_Axis3_ActualPosHiRaw : UINT;  (* 未割付・不使用 IN25 3軸目 現在位置 上位 [0.01mm] *)
    RCON2_IN_Axis3_CurrentLoRaw : UINT;  (* 未割付・不使用 IN26 3軸目 指令電流 下位 [mA] *)
    RCON2_IN_Axis3_CurrentHiRaw : UINT;  (* 未割付・不使用 IN27 3軸目 指令電流 上位 [mA] *)
    RCON2_IN_Axis3_ActualSpeedRaw : UINT;  (* 未割付・不使用 IN28 3軸目 現在速度 [実機単位・符号付き] *)
    RCON2_IN_Axis3_ReservedInRaw : UINT;  (* 未割付・不使用 IN29 3軸目 予約（使用禁止） *)
    RCON2_IN_Axis3_AlarmCodeRaw : UINT;  (* 未割付・不使用 IN30 3軸目 軸異常コード *)
    RCON2_IN_Axis3_StatusRaw : UINT;  (* 未割付・不使用 IN31 3軸目 状態信号（PEND/SV等） *)
    RCON2_IN_Axis4_ActualPosLoRaw : UINT;  (* 未割付・不使用 IN32 4軸目 現在位置 下位 [0.01mm] *)
    RCON2_IN_Axis4_ActualPosHiRaw : UINT;  (* 未割付・不使用 IN33 4軸目 現在位置 上位 [0.01mm] *)
    RCON2_IN_Axis4_CurrentLoRaw : UINT;  (* 未割付・不使用 IN34 4軸目 指令電流 下位 [mA] *)
    RCON2_IN_Axis4_CurrentHiRaw : UINT;  (* 未割付・不使用 IN35 4軸目 指令電流 上位 [mA] *)
    RCON2_IN_Axis4_ActualSpeedRaw : UINT;  (* 未割付・不使用 IN36 4軸目 現在速度 [実機単位・符号付き] *)
    RCON2_IN_Axis4_ReservedInRaw : UINT;  (* 未割付・不使用 IN37 4軸目 予約（使用禁止） *)
    RCON2_IN_Axis4_AlarmCodeRaw : UINT;  (* 未割付・不使用 IN38 4軸目 軸異常コード *)
    RCON2_IN_Axis4_StatusRaw : UINT;  (* 未割付・不使用 IN39 4軸目 状態信号（PEND/SV等） *)
    RCON2_IN_Axis5_ActualPosLoRaw : UINT;  (* 未割付・不使用 IN40 5軸目 現在位置 下位 [0.01mm] *)
    RCON2_IN_Axis5_ActualPosHiRaw : UINT;  (* 未割付・不使用 IN41 5軸目 現在位置 上位 [0.01mm] *)
    RCON2_IN_Axis5_CurrentLoRaw : UINT;  (* 未割付・不使用 IN42 5軸目 指令電流 下位 [mA] *)
    RCON2_IN_Axis5_CurrentHiRaw : UINT;  (* 未割付・不使用 IN43 5軸目 指令電流 上位 [mA] *)
    RCON2_IN_Axis5_ActualSpeedRaw : UINT;  (* 未割付・不使用 IN44 5軸目 現在速度 [実機単位・符号付き] *)
    RCON2_IN_Axis5_ReservedInRaw : UINT;  (* 未割付・不使用 IN45 5軸目 予約（使用禁止） *)
    RCON2_IN_Axis5_AlarmCodeRaw : UINT;  (* 未割付・不使用 IN46 5軸目 軸異常コード *)
    RCON2_IN_Axis5_StatusRaw : UINT;  (* 未割付・不使用 IN47 5軸目 状態信号（PEND/SV等） *)
    E005_Out_OUT00_2003_01 : UINT;  (* 旧I/O候補（未割付・不使用） *)
    E005_Out_OUT01_2003_02 : UINT;  (* 旧I/O候補（未割付・不使用） *)
    E005_Out_OUT02_2003_03 : UINT;  (* 旧I/O候補（未割付・不使用） *)
    E005_Out_OUT03_2003_04 : UINT;  (* 旧I/O候補（未割付・不使用） *)
    E005_Out_OUT04_2003_05 : UINT;  (* 旧I/O候補（未割付・不使用） *)
    E005_Out_OUT05_2003_06 : UINT;  (* 旧I/O候補（未割付・不使用） *)
    E005_Out_OUT06_2003_07 : UINT;  (* 旧I/O候補（未割付・不使用） *)
    E005_Out_OUT07_2003_08 : UINT;  (* 旧I/O候補（未割付・不使用） *)
    E005_Out_OUT08_2003_09 : UINT;  (* 旧I/O候補（未割付・不使用） *)
    E005_Out_OUT09_2003_0A : UINT;  (* 旧I/O候補（未割付・不使用） *)
    E005_Out_OUT10_2003_0B : UINT;  (* 旧I/O候補（未割付・不使用） *)
    E005_Out_OUT11_2003_0C : UINT;  (* 旧I/O候補（未割付・不使用） *)
    E005_Out_OUT12_2003_0D : UINT;  (* 旧I/O候補（未割付・不使用） *)
    E005_Out_OUT13_2003_0E : UINT;  (* 旧I/O候補（未割付・不使用） *)
    E005_Out_OUT14_2003_0F : UINT;  (* 旧I/O候補（未割付・不使用） *)
    E005_Out_OUT15_2003_10 : UINT;  (* 旧I/O候補（未割付・不使用） *)
    E005_Out_OUT16_2003_11 : UINT;  (* 旧I/O候補（未割付・不使用） *)
    E005_Out_OUT17_2003_12 : UINT;  (* 旧I/O候補（未割付・不使用） *)
    E005_Out_OUT18_2003_13 : UINT;  (* 旧I/O候補（未割付・不使用） *)
    E005_Out_OUT19_2003_14 : UINT;  (* 旧I/O候補（未割付・不使用） *)
    E005_Out_OUT20_2003_15 : UINT;  (* 旧I/O候補（未割付・不使用） *)
    E005_Out_OUT21_2003_16 : UINT;  (* 旧I/O候補（未割付・不使用） *)
    E005_Out_OUT22_2003_17 : UINT;  (* 旧I/O候補（未割付・不使用） *)
    E005_Out_OUT23_2003_18 : UINT;  (* 旧I/O候補（未割付・不使用） *)
    E005_Out_OUT24_2003_19 : UINT;  (* 旧I/O候補（未割付・不使用） *)
    E005_Out_OUT25_2003_1A : UINT;  (* 旧I/O候補（未割付・不使用） *)
    E005_Out_OUT26_2003_1B : UINT;  (* 旧I/O候補（未割付・不使用） *)
    E005_Out_OUT27_2003_1C : UINT;  (* 旧I/O候補（未割付・不使用） *)
    E005_Out_OUT28_2003_1D : UINT;  (* 旧I/O候補（未割付・不使用） *)
    E005_Out_OUT29_2003_1E : UINT;  (* 旧I/O候補（未割付・不使用） *)
    E005_Out_OUT30_2003_1F : UINT;  (* 旧I/O候補（未割付・不使用） *)
    E005_Out_OUT31_2003_20 : UINT;  (* 旧I/O候補（未割付・不使用） *)
    E005_Out_OUT32_2003_21 : UINT;  (* 旧I/O候補（未割付・不使用） *)
    E005_Out_OUT33_2003_22 : UINT;  (* 旧I/O候補（未割付・不使用） *)
    E005_Out_OUT34_2003_23 : UINT;  (* 旧I/O候補（未割付・不使用） *)
    E005_Out_OUT35_2003_24 : UINT;  (* 旧I/O候補（未割付・不使用） *)
    E005_Out_OUT36_2003_25 : UINT;  (* 旧I/O候補（未割付・不使用） *)
    E005_Out_OUT37_2003_26 : UINT;  (* 旧I/O候補（未割付・不使用） *)
    E005_Out_OUT38_2003_27 : UINT;  (* 旧I/O候補（未割付・不使用） *)
    E005_Out_OUT39_2003_28 : UINT;  (* 旧I/O候補（未割付・不使用） *)
    E005_Out_OUT40_2003_29 : UINT;  (* 旧I/O候補（未割付・不使用） *)
    E005_Out_OUT41_2003_2A : UINT;  (* 旧I/O候補（未割付・不使用） *)
    E005_Out_OUT42_2003_2B : UINT;  (* 旧I/O候補（未割付・不使用） *)
    E005_Out_OUT43_2003_2C : UINT;  (* 旧I/O候補（未割付・不使用） *)
    E005_Out_OUT44_2003_2D : UINT;  (* 旧I/O候補（未割付・不使用） *)
    E005_Out_OUT45_2003_2E : UINT;  (* 旧I/O候補（未割付・不使用） *)
    E005_Out_OUT46_2003_2F : UINT;  (* 旧I/O候補（未割付・不使用） *)
    E005_Out_OUT47_2003_30 : UINT;  (* 旧I/O候補（未割付・不使用） *)
    E005_Out_OUT48_2003_31 : UINT;  (* 旧I/O候補（未割付・不使用） *)
    E005_Out_OUT49_2003_32 : UINT;  (* 旧I/O候補（未割付・不使用） *)
    E005_Out_OUT50_2003_33 : UINT;  (* 旧I/O候補（未割付・不使用） *)
    E005_Out_OUT51_2003_34 : UINT;  (* 旧I/O候補（未割付・不使用） *)
    E005_Out_OUT52_2003_35 : UINT;  (* 旧I/O候補（未割付・不使用） *)
    E005_Out_OUT53_2003_36 : UINT;  (* 旧I/O候補（未割付・不使用） *)
    E005_Out_OUT54_2003_37 : UINT;  (* 旧I/O候補（未割付・不使用） *)
    E005_Out_OUT55_2003_38 : UINT;  (* 旧I/O候補（未割付・不使用） *)
    E005_Out_OUT56_2003_39 : UINT;  (* 旧I/O候補（未割付・不使用） *)
    E005_Out_OUT57_2003_3A : UINT;  (* 旧I/O候補（未割付・不使用） *)
    E005_Out_OUT58_2003_3B : UINT;  (* 旧I/O候補（未割付・不使用） *)
    E005_Out_OUT59_2003_3C : UINT;  (* 旧I/O候補（未割付・不使用） *)
    E005_Out_OUT60_2003_3D : UINT;  (* 旧I/O候補（未割付・不使用） *)
    E005_Out_OUT61_2003_3E : UINT;  (* 旧I/O候補（未割付・不使用） *)
    E005_Out_OUT62_2003_3F : UINT;  (* 旧I/O候補（未割付・不使用） *)
    E005_Out_OUT63_2003_40 : UINT;  (* 旧I/O候補（未割付・不使用） *)
    E005_Out_OUT64_2003_41 : UINT;  (* 旧I/O候補（未割付・不使用） *)
    E005_Out_OUT65_2003_42 : UINT;  (* 旧I/O候補（未割付・不使用） *)
    E005_Out_OUT66_2003_43 : UINT;  (* 旧I/O候補（未割付・不使用） *)
    E005_Out_OUT67_2003_44 : UINT;  (* 旧I/O候補（未割付・不使用） *)
    E005_Out_OUT68_2003_45 : UINT;  (* 旧I/O候補（未割付・不使用） *)
    E005_Out_OUT69_2003_46 : UINT;  (* 旧I/O候補（未割付・不使用） *)
    E005_Out_OUT70_2003_47 : UINT;  (* 旧I/O候補（未割付・不使用） *)
    E005_Out_OUT71_2003_48 : UINT;  (* 旧I/O候補（未割付・不使用） *)
    E005_In_IN00_2004_01 : UINT;  (* 旧I/O候補（未割付・不使用） *)
    E005_In_IN01_2004_02 : UINT;  (* 旧I/O候補（未割付・不使用） *)
    E005_In_IN02_2004_03 : UINT;  (* 旧I/O候補（未割付・不使用） *)
    E005_In_IN03_2004_04 : UINT;  (* 旧I/O候補（未割付・不使用） *)
    E005_In_IN04_2004_05 : UINT;  (* 旧I/O候補（未割付・不使用） *)
    E005_In_IN05_2004_06 : UINT;  (* 旧I/O候補（未割付・不使用） *)
    E005_In_IN06_2004_07 : UINT;  (* 旧I/O候補（未割付・不使用） *)
    E005_In_IN07_2004_08 : UINT;  (* 旧I/O候補（未割付・不使用） *)
    E005_In_IN08_2004_09 : UINT;  (* 旧I/O候補（未割付・不使用） *)
    E005_In_IN09_2004_0A : UINT;  (* 旧I/O候補（未割付・不使用） *)
    E005_In_IN10_2004_0B : UINT;  (* 旧I/O候補（未割付・不使用） *)
    E005_In_IN11_2004_0C : UINT;  (* 旧I/O候補（未割付・不使用） *)
    E005_In_IN12_2004_0D : UINT;  (* 旧I/O候補（未割付・不使用） *)
    E005_In_IN13_2004_0E : UINT;  (* 旧I/O候補（未割付・不使用） *)
    E005_In_IN14_2004_0F : UINT;  (* 旧I/O候補（未割付・不使用） *)
    E005_In_IN15_2004_10 : UINT;  (* 旧I/O候補（未割付・不使用） *)
    E005_In_IN16_2004_11 : UINT;  (* 旧I/O候補（未割付・不使用） *)
    E005_In_IN17_2004_12 : UINT;  (* 旧I/O候補（未割付・不使用） *)
    E005_In_IN18_2004_13 : UINT;  (* 旧I/O候補（未割付・不使用） *)
    E005_In_IN19_2004_14 : UINT;  (* 旧I/O候補（未割付・不使用） *)
    E005_In_IN20_2004_15 : UINT;  (* 旧I/O候補（未割付・不使用） *)
    E005_In_IN21_2004_16 : UINT;  (* 旧I/O候補（未割付・不使用） *)
    E005_In_IN22_2004_17 : UINT;  (* 旧I/O候補（未割付・不使用） *)
    E005_In_IN23_2004_18 : UINT;  (* 旧I/O候補（未割付・不使用） *)
    E005_In_IN24_2004_19 : UINT;  (* 旧I/O候補（未割付・不使用） *)
    E005_In_IN25_2004_1A : UINT;  (* 旧I/O候補（未割付・不使用） *)
    E005_In_IN26_2004_1B : UINT;  (* 旧I/O候補（未割付・不使用） *)
    E005_In_IN27_2004_1C : UINT;  (* 旧I/O候補（未割付・不使用） *)
    E005_In_IN28_2004_1D : UINT;  (* 旧I/O候補（未割付・不使用） *)
    E005_In_IN29_2004_1E : UINT;  (* 旧I/O候補（未割付・不使用） *)
    E005_In_IN30_2004_1F : UINT;  (* 旧I/O候補（未割付・不使用） *)
    E005_In_IN31_2004_20 : UINT;  (* 旧I/O候補（未割付・不使用） *)
    E005_In_IN32_2004_21 : UINT;  (* 旧I/O候補（未割付・不使用） *)
    E005_In_IN33_2004_22 : UINT;  (* 旧I/O候補（未割付・不使用） *)
    E005_In_IN34_2004_23 : UINT;  (* 旧I/O候補（未割付・不使用） *)
    E005_In_IN35_2004_24 : UINT;  (* 旧I/O候補（未割付・不使用） *)
    E005_In_IN36_2004_25 : UINT;  (* 旧I/O候補（未割付・不使用） *)
    E005_In_IN37_2004_26 : UINT;  (* 旧I/O候補（未割付・不使用） *)
    E005_In_IN38_2004_27 : UINT;  (* 旧I/O候補（未割付・不使用） *)
    E005_In_IN39_2004_28 : UINT;  (* 旧I/O候補（未割付・不使用） *)
    E005_In_IN40_2004_29 : UINT;  (* 旧I/O候補（未割付・不使用） *)
    E005_In_IN41_2004_2A : UINT;  (* 旧I/O候補（未割付・不使用） *)
    E005_In_IN42_2004_2B : UINT;  (* 旧I/O候補（未割付・不使用） *)
    E005_In_IN43_2004_2C : UINT;  (* 旧I/O候補（未割付・不使用） *)
    E005_In_IN44_2004_2D : UINT;  (* 旧I/O候補（未割付・不使用） *)
    E005_In_IN45_2004_2E : UINT;  (* 旧I/O候補（未割付・不使用） *)
    E005_In_IN46_2004_2F : UINT;  (* 旧I/O候補（未割付・不使用） *)
    E005_In_IN47_2004_30 : UINT;  (* 旧I/O候補（未割付・不使用） *)
    E005_In_IN48_2004_31 : UINT;  (* 旧I/O候補（未割付・不使用） *)
    E005_In_IN49_2004_32 : UINT;  (* 旧I/O候補（未割付・不使用） *)
    E005_In_IN50_2004_33 : UINT;  (* 旧I/O候補（未割付・不使用） *)
    E005_In_IN51_2004_34 : UINT;  (* 旧I/O候補（未割付・不使用） *)
    E005_In_IN52_2004_35 : UINT;  (* 旧I/O候補（未割付・不使用） *)
    E005_In_IN53_2004_36 : UINT;  (* 旧I/O候補（未割付・不使用） *)
    E005_In_IN54_2004_37 : UINT;  (* 旧I/O候補（未割付・不使用） *)
    E005_In_IN55_2004_38 : UINT;  (* 旧I/O候補（未割付・不使用） *)
    E005_In_IN56_2004_39 : UINT;  (* 旧I/O候補（未割付・不使用） *)
    E005_In_IN57_2004_3A : UINT;  (* 旧I/O候補（未割付・不使用） *)
    E005_In_IN58_2004_3B : UINT;  (* 旧I/O候補（未割付・不使用） *)
    E005_In_IN59_2004_3C : UINT;  (* 旧I/O候補（未割付・不使用） *)
    E005_In_IN60_2004_3D : UINT;  (* 旧I/O候補（未割付・不使用） *)
    E005_In_IN61_2004_3E : UINT;  (* 旧I/O候補（未割付・不使用） *)
    E005_In_IN62_2004_3F : UINT;  (* 旧I/O候補（未割付・不使用） *)
    E005_In_IN63_2004_40 : UINT;  (* 旧I/O候補（未割付・不使用） *)
    E005_In_IN64_2004_41 : UINT;  (* 旧I/O候補（未割付・不使用） *)
    E005_In_IN65_2004_42 : UINT;  (* 旧I/O候補（未割付・不使用） *)
    E005_In_IN66_2004_43 : UINT;  (* 旧I/O候補（未割付・不使用） *)
    E005_In_IN67_2004_44 : UINT;  (* 旧I/O候補（未割付・不使用） *)
    E005_In_IN68_2004_45 : UINT;  (* 旧I/O候補（未割付・不使用） *)
    E005_In_IN69_2004_46 : UINT;  (* 旧I/O候補（未割付・不使用） *)
    E005_In_IN70_2004_47 : UINT;  (* 旧I/O候補（未割付・不使用） *)
    E005_In_IN71_2004_48 : UINT;  (* 旧I/O候補（未割付・不使用） *)
    E005_Out_OUT00_2003_01_1 : UINT;  (* OUT00 共通制御（MON/RTE）; at ECAT://node#5/Out_OUT00_2003_01 *)
    E005_Out_OUT01_2003_02_1 : UINT;  (* OUT01 予約（書込禁止）; at ECAT://node#5/Out_OUT01_2003_02 *)
    E005_Out_OUT02_2003_03_1 : UINT;  (* OUT02 予約（書込禁止）; at ECAT://node#5/Out_OUT02_2003_03 *)
    E005_Out_OUT03_2003_04_1 : UINT;  (* OUT03 予約（書込禁止）; at ECAT://node#5/Out_OUT03_2003_04 *)
    E005_Out_OUT04_2003_05_1 : UINT;  (* OUT04 予約（書込禁止）; at ECAT://node#5/Out_OUT04_2003_05 *)
    E005_Out_OUT05_2003_06_1 : UINT;  (* OUT05 予約（書込禁止）; at ECAT://node#5/Out_OUT05_2003_06 *)
    E005_Out_OUT06_2003_07_1 : UINT;  (* OUT06 予約（書込禁止）; at ECAT://node#5/Out_OUT06_2003_07 *)
    E005_Out_OUT07_2003_08_1 : UINT;  (* OUT07 予約（書込禁止）; at ECAT://node#5/Out_OUT07_2003_08 *)
    E005_Out_OUT08_2003_09_1 : UINT;  (* OUT08 1軸目 目標位置 下位 [0.01mm]; at ECAT://node#5/Out_OUT08_2003_09 *)
    E005_Out_OUT09_2003_0A_1 : UINT;  (* OUT09 1軸目 目標位置 上位 [0.01mm]; at ECAT://node#5/Out_OUT09_2003_0A *)
    E005_Out_OUT10_2003_0B_1 : UINT;  (* OUT10 1軸目 位置決め幅 下位 [0.01mm]; at ECAT://node#5/Out_OUT10_2003_0B *)
    E005_Out_OUT11_2003_0C_1 : UINT;  (* OUT11 1軸目 位置決め幅 上位 [0.01mm]; at ECAT://node#5/Out_OUT11_2003_0C *)
    E005_Out_OUT12_2003_0D_1 : UINT;  (* OUT12 1軸目 速度指令 [実機単位]; at ECAT://node#5/Out_OUT12_2003_0D *)
    E005_Out_OUT13_2003_0E_1 : UINT;  (* OUT13 1軸目 共通加減速 [0.01G]; at ECAT://node#5/Out_OUT13_2003_0E *)
    E005_Out_OUT14_2003_0F_1 : UINT;  (* OUT14 1軸目 押付け制限 [255=100%]; at ECAT://node#5/Out_OUT14_2003_0F *)
    E005_Out_OUT15_2003_10_1 : UINT;  (* OUT15 1軸目 制御信号（DSTR/SON等）; at ECAT://node#5/Out_OUT15_2003_10 *)
    E005_Out_OUT16_2003_11_1 : UINT;  (* OUT16 2軸目 目標位置 下位 [0.01mm]; at ECAT://node#5/Out_OUT16_2003_11 *)
    E005_Out_OUT17_2003_12_1 : UINT;  (* OUT17 2軸目 目標位置 上位 [0.01mm]; at ECAT://node#5/Out_OUT17_2003_12 *)
    E005_Out_OUT18_2003_13_1 : UINT;  (* OUT18 2軸目 位置決め幅 下位 [0.01mm]; at ECAT://node#5/Out_OUT18_2003_13 *)
    E005_Out_OUT19_2003_14_1 : UINT;  (* OUT19 2軸目 位置決め幅 上位 [0.01mm]; at ECAT://node#5/Out_OUT19_2003_14 *)
    E005_Out_OUT20_2003_15_1 : UINT;  (* OUT20 2軸目 速度指令 [実機単位]; at ECAT://node#5/Out_OUT20_2003_15 *)
    E005_Out_OUT21_2003_16_1 : UINT;  (* OUT21 2軸目 共通加減速 [0.01G]; at ECAT://node#5/Out_OUT21_2003_16 *)
    E005_Out_OUT22_2003_17_1 : UINT;  (* OUT22 2軸目 押付け制限 [255=100%]; at ECAT://node#5/Out_OUT22_2003_17 *)
    E005_Out_OUT23_2003_18_1 : UINT;  (* OUT23 2軸目 制御信号（DSTR/SON等）; at ECAT://node#5/Out_OUT23_2003_18 *)
    E005_Out_OUT24_2003_19_1 : UINT;  (* OUT24 3軸目 目標位置 下位 [0.01mm]; at ECAT://node#5/Out_OUT24_2003_19 *)
    E005_Out_OUT25_2003_1A_1 : UINT;  (* OUT25 3軸目 目標位置 上位 [0.01mm]; at ECAT://node#5/Out_OUT25_2003_1A *)
    E005_Out_OUT26_2003_1B_1 : UINT;  (* OUT26 3軸目 位置決め幅 下位 [0.01mm]; at ECAT://node#5/Out_OUT26_2003_1B *)
    E005_Out_OUT27_2003_1C_1 : UINT;  (* OUT27 3軸目 位置決め幅 上位 [0.01mm]; at ECAT://node#5/Out_OUT27_2003_1C *)
    E005_Out_OUT28_2003_1D_1 : UINT;  (* OUT28 3軸目 速度指令 [実機単位]; at ECAT://node#5/Out_OUT28_2003_1D *)
    E005_Out_OUT29_2003_1E_1 : UINT;  (* OUT29 3軸目 共通加減速 [0.01G]; at ECAT://node#5/Out_OUT29_2003_1E *)
    E005_Out_OUT30_2003_1F_1 : UINT;  (* OUT30 3軸目 押付け制限 [255=100%]; at ECAT://node#5/Out_OUT30_2003_1F *)
    E005_Out_OUT31_2003_20_1 : UINT;  (* OUT31 3軸目 制御信号（DSTR/SON等）; at ECAT://node#5/Out_OUT31_2003_20 *)
    E005_Out_OUT32_2003_21_1 : UINT;  (* OUT32 4軸目 目標位置 下位 [0.01mm]; at ECAT://node#5/Out_OUT32_2003_21 *)
    E005_Out_OUT33_2003_22_1 : UINT;  (* OUT33 4軸目 目標位置 上位 [0.01mm]; at ECAT://node#5/Out_OUT33_2003_22 *)
    E005_Out_OUT34_2003_23_1 : UINT;  (* OUT34 4軸目 位置決め幅 下位 [0.01mm]; at ECAT://node#5/Out_OUT34_2003_23 *)
    E005_Out_OUT35_2003_24_1 : UINT;  (* OUT35 4軸目 位置決め幅 上位 [0.01mm]; at ECAT://node#5/Out_OUT35_2003_24 *)
    E005_Out_OUT36_2003_25_1 : UINT;  (* OUT36 4軸目 速度指令 [実機単位]; at ECAT://node#5/Out_OUT36_2003_25 *)
    E005_Out_OUT37_2003_26_1 : UINT;  (* OUT37 4軸目 共通加減速 [0.01G]; at ECAT://node#5/Out_OUT37_2003_26 *)
    E005_Out_OUT38_2003_27_1 : UINT;  (* OUT38 4軸目 押付け制限 [255=100%]; at ECAT://node#5/Out_OUT38_2003_27 *)
    E005_Out_OUT39_2003_28_1 : UINT;  (* OUT39 4軸目 制御信号（DSTR/SON等）; at ECAT://node#5/Out_OUT39_2003_28 *)
    E005_Out_OUT40_2003_29_1 : UINT;  (* OUT40 5軸目 目標位置 下位 [0.01mm]; at ECAT://node#5/Out_OUT40_2003_29 *)
    E005_Out_OUT41_2003_2A_1 : UINT;  (* OUT41 5軸目 目標位置 上位 [0.01mm]; at ECAT://node#5/Out_OUT41_2003_2A *)
    E005_Out_OUT42_2003_2B_1 : UINT;  (* OUT42 5軸目 位置決め幅 下位 [0.01mm]; at ECAT://node#5/Out_OUT42_2003_2B *)
    E005_Out_OUT43_2003_2C_1 : UINT;  (* OUT43 5軸目 位置決め幅 上位 [0.01mm]; at ECAT://node#5/Out_OUT43_2003_2C *)
    E005_Out_OUT44_2003_2D_1 : UINT;  (* OUT44 5軸目 速度指令 [実機単位]; at ECAT://node#5/Out_OUT44_2003_2D *)
    E005_Out_OUT45_2003_2E_1 : UINT;  (* OUT45 5軸目 共通加減速 [0.01G]; at ECAT://node#5/Out_OUT45_2003_2E *)
    E005_Out_OUT46_2003_2F_1 : UINT;  (* OUT46 5軸目 押付け制限 [255=100%]; at ECAT://node#5/Out_OUT46_2003_2F *)
    E005_Out_OUT47_2003_30_1 : UINT;  (* OUT47 5軸目 制御信号（DSTR/SON等）; at ECAT://node#5/Out_OUT47_2003_30 *)
    E005_Out_OUT48_2003_31_1 : UINT;  (* OUT48 用途未確認（今回未使用）; at ECAT://node#5/Out_OUT48_2003_31 *)
    E005_Out_OUT49_2003_32_1 : UINT;  (* OUT49 用途未確認（今回未使用）; at ECAT://node#5/Out_OUT49_2003_32 *)
    E005_Out_OUT50_2003_33_1 : UINT;  (* OUT50 用途未確認（今回未使用）; at ECAT://node#5/Out_OUT50_2003_33 *)
    E005_Out_OUT51_2003_34_1 : UINT;  (* OUT51 用途未確認（今回未使用）; at ECAT://node#5/Out_OUT51_2003_34 *)
    E005_Out_OUT52_2003_35_1 : UINT;  (* OUT52 用途未確認（今回未使用）; at ECAT://node#5/Out_OUT52_2003_35 *)
    E005_Out_OUT53_2003_36_1 : UINT;  (* OUT53 用途未確認（今回未使用）; at ECAT://node#5/Out_OUT53_2003_36 *)
    E005_Out_OUT54_2003_37_1 : UINT;  (* OUT54 用途未確認（今回未使用）; at ECAT://node#5/Out_OUT54_2003_37 *)
    E005_Out_OUT55_2003_38_1 : UINT;  (* OUT55 用途未確認（今回未使用）; at ECAT://node#5/Out_OUT55_2003_38 *)
    E005_In_IN00_2004_01_1 : UINT;  (* IN00 GW状態; at ECAT://node#5/In_IN00_2004_01 *)
    E005_In_IN01_2004_02_1 : UINT;  (* IN01 軸リンク状態; at ECAT://node#5/In_IN01_2004_02 *)
    E005_In_IN02_2004_03_1 : UINT;  (* IN02 電源状態0; at ECAT://node#5/In_IN02_2004_03 *)
    E005_In_IN03_2004_04_1 : UINT;  (* IN03 電源状態1; at ECAT://node#5/In_IN03_2004_04 *)
    E005_In_IN04_2004_05_1 : UINT;  (* IN04 電源状態2; at ECAT://node#5/In_IN04_2004_05 *)
    E005_In_IN05_2004_06_1 : UINT;  (* IN05 電源状態3; at ECAT://node#5/In_IN05_2004_06 *)
    E005_In_IN06_2004_07_1 : UINT;  (* IN06 電源状態4（構成依存）; at ECAT://node#5/In_IN06_2004_07 *)
    E005_In_IN07_2004_08_1 : UINT;  (* IN07 予約（使用禁止）; at ECAT://node#5/In_IN07_2004_08 *)
    E005_In_IN08_2004_09_1 : UINT;  (* IN08 1軸目 現在位置 下位 [0.01mm]; at ECAT://node#5/In_IN08_2004_09 *)
    E005_In_IN09_2004_0A_1 : UINT;  (* IN09 1軸目 現在位置 上位 [0.01mm]; at ECAT://node#5/In_IN09_2004_0A *)
    E005_In_IN10_2004_0B_1 : UINT;  (* IN10 1軸目 指令電流 下位 [mA]; at ECAT://node#5/In_IN10_2004_0B *)
    E005_In_IN11_2004_0C_1 : UINT;  (* IN11 1軸目 指令電流 上位 [mA]; at ECAT://node#5/In_IN11_2004_0C *)
    E005_In_IN12_2004_0D_1 : UINT;  (* IN12 1軸目 現在速度 [実機単位・符号付き]; at ECAT://node#5/In_IN12_2004_0D *)
    E005_In_IN13_2004_0E_1 : UINT;  (* IN13 1軸目 予約（使用禁止）; at ECAT://node#5/In_IN13_2004_0E *)
    E005_In_IN14_2004_0F_1 : UINT;  (* IN14 1軸目 軸異常コード; at ECAT://node#5/In_IN14_2004_0F *)
    E005_In_IN15_2004_10_1 : UINT;  (* IN15 1軸目 状態信号（PEND/SV等）; at ECAT://node#5/In_IN15_2004_10 *)
    E005_In_IN16_2004_11_1 : UINT;  (* IN16 2軸目 現在位置 下位 [0.01mm]; at ECAT://node#5/In_IN16_2004_11 *)
    E005_In_IN17_2004_12_1 : UINT;  (* IN17 2軸目 現在位置 上位 [0.01mm]; at ECAT://node#5/In_IN17_2004_12 *)
    E005_In_IN18_2004_13_1 : UINT;  (* IN18 2軸目 指令電流 下位 [mA]; at ECAT://node#5/In_IN18_2004_13 *)
    E005_In_IN19_2004_14_1 : UINT;  (* IN19 2軸目 指令電流 上位 [mA]; at ECAT://node#5/In_IN19_2004_14 *)
    E005_In_IN20_2004_15_1 : UINT;  (* IN20 2軸目 現在速度 [実機単位・符号付き]; at ECAT://node#5/In_IN20_2004_15 *)
    E005_In_IN21_2004_16_1 : UINT;  (* IN21 2軸目 予約（使用禁止）; at ECAT://node#5/In_IN21_2004_16 *)
    E005_In_IN22_2004_17_1 : UINT;  (* IN22 2軸目 軸異常コード; at ECAT://node#5/In_IN22_2004_17 *)
    E005_In_IN23_2004_18_1 : UINT;  (* IN23 2軸目 状態信号（PEND/SV等）; at ECAT://node#5/In_IN23_2004_18 *)
    E005_In_IN24_2004_19_1 : UINT;  (* IN24 3軸目 現在位置 下位 [0.01mm]; at ECAT://node#5/In_IN24_2004_19 *)
    E005_In_IN25_2004_1A_1 : UINT;  (* IN25 3軸目 現在位置 上位 [0.01mm]; at ECAT://node#5/In_IN25_2004_1A *)
    E005_In_IN26_2004_1B_1 : UINT;  (* IN26 3軸目 指令電流 下位 [mA]; at ECAT://node#5/In_IN26_2004_1B *)
    E005_In_IN27_2004_1C_1 : UINT;  (* IN27 3軸目 指令電流 上位 [mA]; at ECAT://node#5/In_IN27_2004_1C *)
    E005_In_IN28_2004_1D_1 : UINT;  (* IN28 3軸目 現在速度 [実機単位・符号付き]; at ECAT://node#5/In_IN28_2004_1D *)
    E005_In_IN29_2004_1E_1 : UINT;  (* IN29 3軸目 予約（使用禁止）; at ECAT://node#5/In_IN29_2004_1E *)
    E005_In_IN30_2004_1F_1 : UINT;  (* IN30 3軸目 軸異常コード; at ECAT://node#5/In_IN30_2004_1F *)
    E005_In_IN31_2004_20_1 : UINT;  (* IN31 3軸目 状態信号（PEND/SV等）; at ECAT://node#5/In_IN31_2004_20 *)
    E005_In_IN32_2004_21_1 : UINT;  (* IN32 4軸目 現在位置 下位 [0.01mm]; at ECAT://node#5/In_IN32_2004_21 *)
    E005_In_IN33_2004_22_1 : UINT;  (* IN33 4軸目 現在位置 上位 [0.01mm]; at ECAT://node#5/In_IN33_2004_22 *)
    E005_In_IN34_2004_23_1 : UINT;  (* IN34 4軸目 指令電流 下位 [mA]; at ECAT://node#5/In_IN34_2004_23 *)
    E005_In_IN35_2004_24_1 : UINT;  (* IN35 4軸目 指令電流 上位 [mA]; at ECAT://node#5/In_IN35_2004_24 *)
    E005_In_IN36_2004_25_1 : UINT;  (* IN36 4軸目 現在速度 [実機単位・符号付き]; at ECAT://node#5/In_IN36_2004_25 *)
    E005_In_IN37_2004_26_1 : UINT;  (* IN37 4軸目 予約（使用禁止）; at ECAT://node#5/In_IN37_2004_26 *)
    E005_In_IN38_2004_27_1 : UINT;  (* IN38 4軸目 軸異常コード; at ECAT://node#5/In_IN38_2004_27 *)
    E005_In_IN39_2004_28_1 : UINT;  (* IN39 4軸目 状態信号（PEND/SV等）; at ECAT://node#5/In_IN39_2004_28 *)
    E005_In_IN40_2004_29_1 : UINT;  (* IN40 5軸目 現在位置 下位 [0.01mm]; at ECAT://node#5/In_IN40_2004_29 *)
    E005_In_IN41_2004_2A_1 : UINT;  (* IN41 5軸目 現在位置 上位 [0.01mm]; at ECAT://node#5/In_IN41_2004_2A *)
    E005_In_IN42_2004_2B_1 : UINT;  (* IN42 5軸目 指令電流 下位 [mA]; at ECAT://node#5/In_IN42_2004_2B *)
    E005_In_IN43_2004_2C_1 : UINT;  (* IN43 5軸目 指令電流 上位 [mA]; at ECAT://node#5/In_IN43_2004_2C *)
    E005_In_IN44_2004_2D_1 : UINT;  (* IN44 5軸目 現在速度 [実機単位・符号付き]; at ECAT://node#5/In_IN44_2004_2D *)
    E005_In_IN45_2004_2E_1 : UINT;  (* IN45 5軸目 予約（使用禁止）; at ECAT://node#5/In_IN45_2004_2E *)
    E005_In_IN46_2004_2F_1 : UINT;  (* IN46 5軸目 軸異常コード; at ECAT://node#5/In_IN46_2004_2F *)
    E005_In_IN47_2004_30_1 : UINT;  (* IN47 5軸目 状態信号（PEND/SV等）; at ECAT://node#5/In_IN47_2004_30 *)
    E005_In_IN48_2004_31_1 : UINT;  (* IN48 用途未確認（今回未使用）; at ECAT://node#5/In_IN48_2004_31 *)
    E005_In_IN49_2004_32_1 : UINT;  (* IN49 用途未確認（今回未使用）; at ECAT://node#5/In_IN49_2004_32 *)
    E005_In_IN50_2004_33_1 : UINT;  (* IN50 用途未確認（今回未使用）; at ECAT://node#5/In_IN50_2004_33 *)
    E005_In_IN51_2004_34_1 : UINT;  (* IN51 用途未確認（今回未使用）; at ECAT://node#5/In_IN51_2004_34 *)
    E005_In_IN52_2004_35_1 : UINT;  (* IN52 用途未確認（今回未使用）; at ECAT://node#5/In_IN52_2004_35 *)
    E005_In_IN53_2004_36_1 : UINT;  (* IN53 用途未確認（今回未使用）; at ECAT://node#5/In_IN53_2004_36 *)
    E005_In_IN54_2004_37_1 : UINT;  (* IN54 用途未確認（今回未使用）; at ECAT://node#5/In_IN54_2004_37 *)
    E005_In_IN55_2004_38_1 : UINT;  (* IN55 用途未確認（今回未使用）; at ECAT://node#5/In_IN55_2004_38 *)
    E001_Out_OUT00_2003_01 : UINT;  (* OUT00 共通制御（MON/RTE）; at ECAT://node#1/Out_OUT00_2003_01 *)
    E001_Out_OUT01_2003_02 : UINT;  (* OUT01 予約（書込禁止）; at ECAT://node#1/Out_OUT01_2003_02 *)
    E001_Out_OUT02_2003_03 : UINT;  (* OUT02 予約（書込禁止）; at ECAT://node#1/Out_OUT02_2003_03 *)
    E001_Out_OUT03_2003_04 : UINT;  (* OUT03 予約（書込禁止）; at ECAT://node#1/Out_OUT03_2003_04 *)
    E001_Out_OUT04_2003_05 : UINT;  (* OUT04 予約（書込禁止）; at ECAT://node#1/Out_OUT04_2003_05 *)
    E001_Out_OUT05_2003_06 : UINT;  (* OUT05 予約（書込禁止）; at ECAT://node#1/Out_OUT05_2003_06 *)
    E001_Out_OUT06_2003_07 : UINT;  (* OUT06 予約（書込禁止）; at ECAT://node#1/Out_OUT06_2003_07 *)
    E001_Out_OUT07_2003_08 : UINT;  (* OUT07 予約（書込禁止）; at ECAT://node#1/Out_OUT07_2003_08 *)
    E001_Out_OUT08_2003_09 : UINT;  (* OUT08 目標位置 下位 [0.01mm]; at ECAT://node#1/Out_OUT08_2003_09 *)
    E001_Out_OUT09_2003_0A : UINT;  (* OUT09 目標位置 上位 [0.01mm]; at ECAT://node#1/Out_OUT09_2003_0A *)
    E001_Out_OUT10_2003_0B : UINT;  (* OUT10 位置決め幅 下位 [0.01mm]; at ECAT://node#1/Out_OUT10_2003_0B *)
    E001_Out_OUT11_2003_0C : UINT;  (* OUT11 位置決め幅 上位 [0.01mm]; at ECAT://node#1/Out_OUT11_2003_0C *)
    E001_Out_OUT12_2003_0D : UINT;  (* OUT12 速度指令 [実機単位]; at ECAT://node#1/Out_OUT12_2003_0D *)
    E001_Out_OUT13_2003_0E : UINT;  (* OUT13 共通加減速 [0.01G]; at ECAT://node#1/Out_OUT13_2003_0E *)
    E001_Out_OUT14_2003_0F : UINT;  (* OUT14 押付け制限 [255=100%]; at ECAT://node#1/Out_OUT14_2003_0F *)
    E001_Out_OUT15_2003_10 : UINT;  (* OUT15 制御信号（DSTR/SON等）; at ECAT://node#1/Out_OUT15_2003_10 *)
    E001_Out_OUT16_2003_11 : UINT;  (* OUT16 目標位置 下位 [0.01mm]; at ECAT://node#1/Out_OUT16_2003_11 *)
    E001_Out_OUT17_2003_12 : UINT;  (* OUT17 目標位置 上位 [0.01mm]; at ECAT://node#1/Out_OUT17_2003_12 *)
    E001_Out_OUT18_2003_13 : UINT;  (* OUT18 位置決め幅 下位 [0.01mm]; at ECAT://node#1/Out_OUT18_2003_13 *)
    E001_Out_OUT19_2003_14 : UINT;  (* OUT19 位置決め幅 上位 [0.01mm]; at ECAT://node#1/Out_OUT19_2003_14 *)
    E001_Out_OUT20_2003_15 : UINT;  (* OUT20 速度指令 [実機単位]; at ECAT://node#1/Out_OUT20_2003_15 *)
    E001_Out_OUT21_2003_16 : UINT;  (* OUT21 共通加減速 [0.01G]; at ECAT://node#1/Out_OUT21_2003_16 *)
    E001_Out_OUT22_2003_17 : UINT;  (* OUT22 押付け制限 [255=100%]; at ECAT://node#1/Out_OUT22_2003_17 *)
    E001_Out_OUT23_2003_18 : UINT;  (* OUT23 制御信号（DSTR/SON等）; at ECAT://node#1/Out_OUT23_2003_18 *)
    E001_Out_OUT24_2003_19 : UINT;  (* OUT24 目標位置 下位 [0.01mm]; at ECAT://node#1/Out_OUT24_2003_19 *)
    E001_Out_OUT25_2003_1A : UINT;  (* OUT25 目標位置 上位 [0.01mm]; at ECAT://node#1/Out_OUT25_2003_1A *)
    E001_Out_OUT26_2003_1B : UINT;  (* OUT26 位置決め幅 下位 [0.01mm]; at ECAT://node#1/Out_OUT26_2003_1B *)
    E001_Out_OUT27_2003_1C : UINT;  (* OUT27 位置決め幅 上位 [0.01mm]; at ECAT://node#1/Out_OUT27_2003_1C *)
    E001_Out_OUT28_2003_1D : UINT;  (* OUT28 速度指令 [実機単位]; at ECAT://node#1/Out_OUT28_2003_1D *)
    E001_Out_OUT29_2003_1E : UINT;  (* OUT29 共通加減速 [0.01G]; at ECAT://node#1/Out_OUT29_2003_1E *)
    E001_Out_OUT30_2003_1F : UINT;  (* OUT30 押付け制限 [255=100%]; at ECAT://node#1/Out_OUT30_2003_1F *)
    E001_Out_OUT31_2003_20 : UINT;  (* OUT31 制御信号（DSTR/SON等）; at ECAT://node#1/Out_OUT31_2003_20 *)
    E001_Out_OUT32_2003_21 : UINT;  (* OUT32 目標位置 下位 [0.01mm]; at ECAT://node#1/Out_OUT32_2003_21 *)
    E001_Out_OUT33_2003_22 : UINT;  (* OUT33 目標位置 上位 [0.01mm]; at ECAT://node#1/Out_OUT33_2003_22 *)
    E001_Out_OUT34_2003_23 : UINT;  (* OUT34 位置決め幅 下位 [0.01mm]; at ECAT://node#1/Out_OUT34_2003_23 *)
    E001_Out_OUT35_2003_24 : UINT;  (* OUT35 位置決め幅 上位 [0.01mm]; at ECAT://node#1/Out_OUT35_2003_24 *)
    E001_Out_OUT36_2003_25 : UINT;  (* OUT36 速度指令 [実機単位]; at ECAT://node#1/Out_OUT36_2003_25 *)
    E001_Out_OUT37_2003_26 : UINT;  (* OUT37 共通加減速 [0.01G]; at ECAT://node#1/Out_OUT37_2003_26 *)
    E001_Out_OUT38_2003_27 : UINT;  (* OUT38 押付け制限 [255=100%]; at ECAT://node#1/Out_OUT38_2003_27 *)
    E001_Out_OUT39_2003_28 : UINT;  (* OUT39 制御信号（DSTR/SON等）; at ECAT://node#1/Out_OUT39_2003_28 *)
    E001_Out_OUT40_2003_29 : UINT;  (* OUT40 目標位置 下位 [0.01mm]; at ECAT://node#1/Out_OUT40_2003_29 *)
    E001_Out_OUT41_2003_2A : UINT;  (* OUT41 目標位置 上位 [0.01mm]; at ECAT://node#1/Out_OUT41_2003_2A *)
    E001_Out_OUT42_2003_2B : UINT;  (* OUT42 位置決め幅 下位 [0.01mm]; at ECAT://node#1/Out_OUT42_2003_2B *)
    E001_Out_OUT43_2003_2C : UINT;  (* OUT43 位置決め幅 上位 [0.01mm]; at ECAT://node#1/Out_OUT43_2003_2C *)
    E001_Out_OUT44_2003_2D : UINT;  (* OUT44 速度指令 [実機単位]; at ECAT://node#1/Out_OUT44_2003_2D *)
    E001_Out_OUT45_2003_2E : UINT;  (* OUT45 共通加減速 [0.01G]; at ECAT://node#1/Out_OUT45_2003_2E *)
    E001_Out_OUT46_2003_2F : UINT;  (* OUT46 押付け制限 [255=100%]; at ECAT://node#1/Out_OUT46_2003_2F *)
    E001_Out_OUT47_2003_30 : UINT;  (* OUT47 制御信号（DSTR/SON等）; at ECAT://node#1/Out_OUT47_2003_30 *)
    E001_Out_OUT48_2003_31 : UINT;  (* OUT48 目標位置 下位 [0.01mm]; at ECAT://node#1/Out_OUT48_2003_31 *)
    E001_Out_OUT49_2003_32 : UINT;  (* OUT49 目標位置 上位 [0.01mm]; at ECAT://node#1/Out_OUT49_2003_32 *)
    E001_Out_OUT50_2003_33 : UINT;  (* OUT50 位置決め幅 下位 [0.01mm]; at ECAT://node#1/Out_OUT50_2003_33 *)
    E001_Out_OUT51_2003_34 : UINT;  (* OUT51 位置決め幅 上位 [0.01mm]; at ECAT://node#1/Out_OUT51_2003_34 *)
    E001_Out_OUT52_2003_35 : UINT;  (* OUT52 速度指令 [実機単位]; at ECAT://node#1/Out_OUT52_2003_35 *)
    E001_Out_OUT53_2003_36 : UINT;  (* OUT53 共通加減速 [0.01G]; at ECAT://node#1/Out_OUT53_2003_36 *)
    E001_Out_OUT54_2003_37 : UINT;  (* OUT54 押付け制限 [255=100%]; at ECAT://node#1/Out_OUT54_2003_37 *)
    E001_Out_OUT55_2003_38 : UINT;  (* OUT55 制御信号（DSTR/SON等）; at ECAT://node#1/Out_OUT55_2003_38 *)
    E001_Out_OUT56_2003_39 : UINT;  (* OUT56 112Byte範囲外（未割付・不使用） *)
    E001_Out_OUT57_2003_3A : UINT;  (* OUT57 112Byte範囲外（未割付・不使用） *)
    E001_Out_OUT58_2003_3B : UINT;  (* OUT58 112Byte範囲外（未割付・不使用） *)
    E001_Out_OUT59_2003_3C : UINT;  (* OUT59 112Byte範囲外（未割付・不使用） *)
    E001_Out_OUT60_2003_3D : UINT;  (* OUT60 112Byte範囲外（未割付・不使用） *)
    E001_Out_OUT61_2003_3E : UINT;  (* OUT61 112Byte範囲外（未割付・不使用） *)
    E001_Out_OUT62_2003_3F : UINT;  (* OUT62 112Byte範囲外（未割付・不使用） *)
    E001_Out_OUT63_2003_40 : UINT;  (* OUT63 112Byte範囲外（未割付・不使用） *)
    E001_Out_OUT64_2003_41 : UINT;  (* OUT64 112Byte範囲外（未割付・不使用） *)
    E001_Out_OUT65_2003_42 : UINT;  (* OUT65 112Byte範囲外（未割付・不使用） *)
    E001_Out_OUT66_2003_43 : UINT;  (* OUT66 112Byte範囲外（未割付・不使用） *)
    E001_Out_OUT67_2003_44 : UINT;  (* OUT67 112Byte範囲外（未割付・不使用） *)
    E001_Out_OUT68_2003_45 : UINT;  (* OUT68 112Byte範囲外（未割付・不使用） *)
    E001_Out_OUT69_2003_46 : UINT;  (* OUT69 112Byte範囲外（未割付・不使用） *)
    E001_Out_OUT70_2003_47 : UINT;  (* OUT70 112Byte範囲外（未割付・不使用） *)
    E001_Out_OUT71_2003_48 : UINT;  (* OUT71 112Byte範囲外（未割付・不使用） *)
    E001_In_IN00_2004_01 : UINT;  (* IN00 GW状態; at ECAT://node#1/In_IN00_2004_01 *)
    E001_In_IN01_2004_02 : UINT;  (* IN01 軸リンク状態; at ECAT://node#1/In_IN01_2004_02 *)
    E001_In_IN02_2004_03 : UINT;  (* IN02 電源状態0; at ECAT://node#1/In_IN02_2004_03 *)
    E001_In_IN03_2004_04 : UINT;  (* IN03 電源状態1; at ECAT://node#1/In_IN03_2004_04 *)
    E001_In_IN04_2004_05 : UINT;  (* IN04 電源状態2; at ECAT://node#1/In_IN04_2004_05 *)
    E001_In_IN05_2004_06 : UINT;  (* IN05 電源状態3; at ECAT://node#1/In_IN05_2004_06 *)
    E001_In_IN06_2004_07 : UINT;  (* IN06 電源状態4（構成依存）; at ECAT://node#1/In_IN06_2004_07 *)
    E001_In_IN07_2004_08 : UINT;  (* IN07 予約（使用禁止）; at ECAT://node#1/In_IN07_2004_08 *)
    E001_In_IN08_2004_09 : UINT;  (* IN08 現在位置 下位 [0.01mm]; at ECAT://node#1/In_IN08_2004_09 *)
    E001_In_IN09_2004_0A : UINT;  (* IN09 現在位置 上位 [0.01mm]; at ECAT://node#1/In_IN09_2004_0A *)
    E001_In_IN10_2004_0B : UINT;  (* IN10 指令電流 下位 [mA]; at ECAT://node#1/In_IN10_2004_0B *)
    E001_In_IN11_2004_0C : UINT;  (* IN11 指令電流 上位 [mA]; at ECAT://node#1/In_IN11_2004_0C *)
    E001_In_IN12_2004_0D : UINT;  (* IN12 現在速度 [実機単位・符号付き]; at ECAT://node#1/In_IN12_2004_0D *)
    E001_In_IN13_2004_0E : UINT;  (* IN13 予約（使用禁止）; at ECAT://node#1/In_IN13_2004_0E *)
    E001_In_IN14_2004_0F : UINT;  (* IN14 軸異常コード; at ECAT://node#1/In_IN14_2004_0F *)
    E001_In_IN15_2004_10 : UINT;  (* IN15 状態信号（PEND/SV等）; at ECAT://node#1/In_IN15_2004_10 *)
    E001_In_IN16_2004_11 : UINT;  (* IN16 現在位置 下位 [0.01mm]; at ECAT://node#1/In_IN16_2004_11 *)
    E001_In_IN17_2004_12 : UINT;  (* IN17 現在位置 上位 [0.01mm]; at ECAT://node#1/In_IN17_2004_12 *)
    E001_In_IN18_2004_13 : UINT;  (* IN18 指令電流 下位 [mA]; at ECAT://node#1/In_IN18_2004_13 *)
    E001_In_IN19_2004_14 : UINT;  (* IN19 指令電流 上位 [mA]; at ECAT://node#1/In_IN19_2004_14 *)
    E001_In_IN20_2004_15 : UINT;  (* IN20 現在速度 [実機単位・符号付き]; at ECAT://node#1/In_IN20_2004_15 *)
    E001_In_IN21_2004_16 : UINT;  (* IN21 予約（使用禁止）; at ECAT://node#1/In_IN21_2004_16 *)
    E001_In_IN22_2004_17 : UINT;  (* IN22 軸異常コード; at ECAT://node#1/In_IN22_2004_17 *)
    E001_In_IN23_2004_18 : UINT;  (* IN23 状態信号（PEND/SV等）; at ECAT://node#1/In_IN23_2004_18 *)
    E001_In_IN24_2004_19 : UINT;  (* IN24 現在位置 下位 [0.01mm]; at ECAT://node#1/In_IN24_2004_19 *)
    E001_In_IN25_2004_1A : UINT;  (* IN25 現在位置 上位 [0.01mm]; at ECAT://node#1/In_IN25_2004_1A *)
    E001_In_IN26_2004_1B : UINT;  (* IN26 指令電流 下位 [mA]; at ECAT://node#1/In_IN26_2004_1B *)
    E001_In_IN27_2004_1C : UINT;  (* IN27 指令電流 上位 [mA]; at ECAT://node#1/In_IN27_2004_1C *)
    E001_In_IN28_2004_1D : UINT;  (* IN28 現在速度 [実機単位・符号付き]; at ECAT://node#1/In_IN28_2004_1D *)
    E001_In_IN29_2004_1E : UINT;  (* IN29 予約（使用禁止）; at ECAT://node#1/In_IN29_2004_1E *)
    E001_In_IN30_2004_1F : UINT;  (* IN30 軸異常コード; at ECAT://node#1/In_IN30_2004_1F *)
    E001_In_IN31_2004_20 : UINT;  (* IN31 状態信号（PEND/SV等）; at ECAT://node#1/In_IN31_2004_20 *)
    E001_In_IN32_2004_21 : UINT;  (* IN32 現在位置 下位 [0.01mm]; at ECAT://node#1/In_IN32_2004_21 *)
    E001_In_IN33_2004_22 : UINT;  (* IN33 現在位置 上位 [0.01mm]; at ECAT://node#1/In_IN33_2004_22 *)
    E001_In_IN34_2004_23 : UINT;  (* IN34 指令電流 下位 [mA]; at ECAT://node#1/In_IN34_2004_23 *)
    E001_In_IN35_2004_24 : UINT;  (* IN35 指令電流 上位 [mA]; at ECAT://node#1/In_IN35_2004_24 *)
    E001_In_IN36_2004_25 : UINT;  (* IN36 現在速度 [実機単位・符号付き]; at ECAT://node#1/In_IN36_2004_25 *)
    E001_In_IN37_2004_26 : UINT;  (* IN37 予約（使用禁止）; at ECAT://node#1/In_IN37_2004_26 *)
    E001_In_IN38_2004_27 : UINT;  (* IN38 軸異常コード; at ECAT://node#1/In_IN38_2004_27 *)
    E001_In_IN39_2004_28 : UINT;  (* IN39 状態信号（PEND/SV等）; at ECAT://node#1/In_IN39_2004_28 *)
    E001_In_IN40_2004_29 : UINT;  (* IN40 現在位置 下位 [0.01mm]; at ECAT://node#1/In_IN40_2004_29 *)
    E001_In_IN41_2004_2A : UINT;  (* IN41 現在位置 上位 [0.01mm]; at ECAT://node#1/In_IN41_2004_2A *)
    E001_In_IN42_2004_2B : UINT;  (* IN42 指令電流 下位 [mA]; at ECAT://node#1/In_IN42_2004_2B *)
    E001_In_IN43_2004_2C : UINT;  (* IN43 指令電流 上位 [mA]; at ECAT://node#1/In_IN43_2004_2C *)
    E001_In_IN44_2004_2D : UINT;  (* IN44 現在速度 [実機単位・符号付き]; at ECAT://node#1/In_IN44_2004_2D *)
    E001_In_IN45_2004_2E : UINT;  (* IN45 予約（使用禁止）; at ECAT://node#1/In_IN45_2004_2E *)
    E001_In_IN46_2004_2F : UINT;  (* IN46 軸異常コード; at ECAT://node#1/In_IN46_2004_2F *)
    E001_In_IN47_2004_30 : UINT;  (* IN47 状態信号（PEND/SV等）; at ECAT://node#1/In_IN47_2004_30 *)
    E001_In_IN48_2004_31 : UINT;  (* IN48 現在位置 下位 [0.01mm]; at ECAT://node#1/In_IN48_2004_31 *)
    E001_In_IN49_2004_32 : UINT;  (* IN49 現在位置 上位 [0.01mm]; at ECAT://node#1/In_IN49_2004_32 *)
    E001_In_IN50_2004_33 : UINT;  (* IN50 指令電流 下位 [mA]; at ECAT://node#1/In_IN50_2004_33 *)
    E001_In_IN51_2004_34 : UINT;  (* IN51 指令電流 上位 [mA]; at ECAT://node#1/In_IN51_2004_34 *)
    E001_In_IN52_2004_35 : UINT;  (* IN52 現在速度 [実機単位・符号付き]; at ECAT://node#1/In_IN52_2004_35 *)
    E001_In_IN53_2004_36 : UINT;  (* IN53 予約（使用禁止）; at ECAT://node#1/In_IN53_2004_36 *)
    E001_In_IN54_2004_37 : UINT;  (* IN54 軸異常コード; at ECAT://node#1/In_IN54_2004_37 *)
    E001_In_IN55_2004_38 : UINT;  (* IN55 状態信号（PEND/SV等）; at ECAT://node#1/In_IN55_2004_38 *)
    E001_In_IN56_2004_39 : UINT;  (* IN56 112Byte範囲外（未割付・不使用） *)
    E001_In_IN57_2004_3A : UINT;  (* IN57 112Byte範囲外（未割付・不使用） *)
    E001_In_IN58_2004_3B : UINT;  (* IN58 112Byte範囲外（未割付・不使用） *)
    E001_In_IN59_2004_3C : UINT;  (* IN59 112Byte範囲外（未割付・不使用） *)
    E001_In_IN60_2004_3D : UINT;  (* IN60 112Byte範囲外（未割付・不使用） *)
    E001_In_IN61_2004_3E : UINT;  (* IN61 112Byte範囲外（未割付・不使用） *)
    E001_In_IN62_2004_3F : UINT;  (* IN62 112Byte範囲外（未割付・不使用） *)
    E001_In_IN63_2004_40 : UINT;  (* IN63 112Byte範囲外（未割付・不使用） *)
    E001_In_IN64_2004_41 : UINT;  (* IN64 112Byte範囲外（未割付・不使用） *)
    E001_In_IN65_2004_42 : UINT;  (* IN65 112Byte範囲外（未割付・不使用） *)
    E001_In_IN66_2004_43 : UINT;  (* IN66 112Byte範囲外（未割付・不使用） *)
    E001_In_IN67_2004_44 : UINT;  (* IN67 112Byte範囲外（未割付・不使用） *)
    E001_In_IN68_2004_45 : UINT;  (* IN68 112Byte範囲外（未割付・不使用） *)
    E001_In_IN69_2004_46 : UINT;  (* IN69 112Byte範囲外（未割付・不使用） *)
    E001_In_IN70_2004_47 : UINT;  (* IN70 112Byte範囲外（未割付・不使用） *)
    E001_In_IN71_2004_48 : UINT;  (* IN71 112Byte範囲外（未割付・不使用） *)
    RCON1_RxRaw : ARRAY[0..55] OF UINT;  (* 受信値（バイト交換前）; [0] IN00 GW状態; [1] IN01 軸リンク状態; [2] IN02 電源状態0; [3] IN03 電源状態1; [4] IN04 電源状態2; [5] IN05 電源状態3; [6] IN06 電源状態4（構成依存）; [7] IN07 予約（使用禁止）; [8] IN08 A(左側) RCON1_1 NG1上下降 現在位置 下位 [0.01mm]; [9] IN09 A(左側) RCON1_1 NG1上下降 現在位置 上位 [0.01mm]; [10] IN10 A(左側) RCON1_1 NG1上下降 指令電流 下位 [mA]; [11] IN11 A(左側) RCON1_1 NG1上下降 指令電流 上位 [mA]; [12] IN12 A(左側) RCON1_1 NG1上下降 現在速度 [実機単位・符号付き]; [13] IN13 A(左側) RCON1_1 NG1上下降 予約（使用禁止）; [14] IN14 A(左側) RCON1_1 NG1上下降 軸異常コード; [15] IN15 A(左側) RCON1_1 NG1上下降 状態信号（PEND/SV等）; [16] IN16 B(右側) RCON1_2 NG1上下降 現在位置 下位 [0.01mm]; [17] IN17 B(右側) RCON1_2 NG1上下降 現在位置 上位 [0.01mm]; [18] IN18 B(右側) RCON1_2 NG1上下降 指令電流 下位 [mA]; [19] IN19 B(右側) RCON1_2 NG1上下降 指令電流 上位 [mA]; [20] IN20 B(右側) RCON1_2 NG1上下降 現在速度 [実機単位・符号付き]; [21] IN21 B(右側) RCON1_2 NG1上下降 予約（使用禁止）; [22] IN22 B(右側) RCON1_2 NG1上下降 軸異常コード; [23] IN23 B(右側) RCON1_2 NG1上下降 状態信号（PEND/SV等）; [24] IN24 A(左側) RCON1_3 SF/NG2仕分け(左右) 現在位置 下位 [0.01mm]; [25] IN25 A(左側) RCON1_3 SF/NG2仕分け(左右) 現在位置 上位 [0.01mm]; [26] IN26 A(左側) RCON1_3 SF/NG2仕分け(左右) 指令電流 下位 [mA]; [27] IN27 A(左側) RCON1_3 SF/NG2仕分け(左右) 指令電流 上位 [mA]; [28] IN28 A(左側) RCON1_3 SF/NG2仕分け(左右) 現在速度 [実機単位・符号付き]; [29] IN29 A(左側) RCON1_3 SF/NG2仕分け(左右) 予約（使用禁止）; [30] IN30 A(左側) RCON1_3 SF/NG2仕分け(左右) 軸異常コード; [31] IN31 A(左側) RCON1_3 SF/NG2仕分け(左右) 状態信号（PEND/SV等）; [32] IN32 B(右側) RCON1_4 SF/NG2送り 現在位置 下位 [0.01mm]; [33] IN33 B(右側) RCON1_4 SF/NG2送り 現在位置 上位 [0.01mm]; [34] IN34 B(右側) RCON1_4 SF/NG2送り 指令電流 下位 [mA]; [35] IN35 B(右側) RCON1_4 SF/NG2送り 指令電流 上位 [mA]; [36] IN36 B(右側) RCON1_4 SF/NG2送り 現在速度 [実機単位・符号付き]; [37] IN37 B(右側) RCON1_4 SF/NG2送り 予約（使用禁止）; [38] IN38 B(右側) RCON1_4 SF/NG2送り 軸異常コード; [39] IN39 B(右側) RCON1_4 SF/NG2送り 状態信号（PEND/SV等）; [40] IN40 A(左側) RCON1_5 SF/NG2上下降 現在位置 下位 [0.01mm]; [41] IN41 A(左側) RCON1_5 SF/NG2上下降 現在位置 上位 [0.01mm]; [42] IN42 A(左側) RCON1_5 SF/NG2上下降 指令電流 下位 [mA]; [43] IN43 A(左側) RCON1_5 SF/NG2上下降 指令電流 上位 [mA]; [44] IN44 A(左側) RCON1_5 SF/NG2上下降 現在速度 [実機単位・符号付き]; [45] IN45 A(左側) RCON1_5 SF/NG2上下降 予約（使用禁止）; [46] IN46 A(左側) RCON1_5 SF/NG2上下降 軸異常コード; [47] IN47 A(左側) RCON1_5 SF/NG2上下降 状態信号（PEND/SV等）; [48] IN48 B(右側) RCON1_6 SF/NG2上下降 現在位置 下位 [0.01mm]; [49] IN49 B(右側) RCON1_6 SF/NG2上下降 現在位置 上位 [0.01mm]; [50] IN50 B(右側) RCON1_6 SF/NG2上下降 指令電流 下位 [mA]; [51] IN51 B(右側) RCON1_6 SF/NG2上下降 指令電流 上位 [mA]; [52] IN52 B(右側) RCON1_6 SF/NG2上下降 現在速度 [実機単位・符号付き]; [53] IN53 B(右側) RCON1_6 SF/NG2上下降 予約（使用禁止）; [54] IN54 B(右側) RCON1_6 SF/NG2上下降 軸異常コード; [55] IN55 B(右側) RCON1_6 SF/NG2上下降 状態信号（PEND/SV等） *)
    RCON1_RxWord : ARRAY[0..55] OF WORD;  (* 受信ワード（正規化後）; [0] IN00 GW状態; [1] IN01 軸リンク状態; [2] IN02 電源状態0; [3] IN03 電源状態1; [4] IN04 電源状態2; [5] IN05 電源状態3; [6] IN06 電源状態4（構成依存）; [7] IN07 予約（使用禁止）; [8] IN08 A(左側) RCON1_1 NG1上下降 現在位置 下位 [0.01mm]; [9] IN09 A(左側) RCON1_1 NG1上下降 現在位置 上位 [0.01mm]; [10] IN10 A(左側) RCON1_1 NG1上下降 指令電流 下位 [mA]; [11] IN11 A(左側) RCON1_1 NG1上下降 指令電流 上位 [mA]; [12] IN12 A(左側) RCON1_1 NG1上下降 現在速度 [実機単位・符号付き]; [13] IN13 A(左側) RCON1_1 NG1上下降 予約（使用禁止）; [14] IN14 A(左側) RCON1_1 NG1上下降 軸異常コード; [15] IN15 A(左側) RCON1_1 NG1上下降 状態信号（PEND/SV等）; [16] IN16 B(右側) RCON1_2 NG1上下降 現在位置 下位 [0.01mm]; [17] IN17 B(右側) RCON1_2 NG1上下降 現在位置 上位 [0.01mm]; [18] IN18 B(右側) RCON1_2 NG1上下降 指令電流 下位 [mA]; [19] IN19 B(右側) RCON1_2 NG1上下降 指令電流 上位 [mA]; [20] IN20 B(右側) RCON1_2 NG1上下降 現在速度 [実機単位・符号付き]; [21] IN21 B(右側) RCON1_2 NG1上下降 予約（使用禁止）; [22] IN22 B(右側) RCON1_2 NG1上下降 軸異常コード; [23] IN23 B(右側) RCON1_2 NG1上下降 状態信号（PEND/SV等）; [24] IN24 A(左側) RCON1_3 SF/NG2仕分け(左右) 現在位置 下位 [0.01mm]; [25] IN25 A(左側) RCON1_3 SF/NG2仕分け(左右) 現在位置 上位 [0.01mm]; [26] IN26 A(左側) RCON1_3 SF/NG2仕分け(左右) 指令電流 下位 [mA]; [27] IN27 A(左側) RCON1_3 SF/NG2仕分け(左右) 指令電流 上位 [mA]; [28] IN28 A(左側) RCON1_3 SF/NG2仕分け(左右) 現在速度 [実機単位・符号付き]; [29] IN29 A(左側) RCON1_3 SF/NG2仕分け(左右) 予約（使用禁止）; [30] IN30 A(左側) RCON1_3 SF/NG2仕分け(左右) 軸異常コード; [31] IN31 A(左側) RCON1_3 SF/NG2仕分け(左右) 状態信号（PEND/SV等）; [32] IN32 B(右側) RCON1_4 SF/NG2送り 現在位置 下位 [0.01mm]; [33] IN33 B(右側) RCON1_4 SF/NG2送り 現在位置 上位 [0.01mm]; [34] IN34 B(右側) RCON1_4 SF/NG2送り 指令電流 下位 [mA]; [35] IN35 B(右側) RCON1_4 SF/NG2送り 指令電流 上位 [mA]; [36] IN36 B(右側) RCON1_4 SF/NG2送り 現在速度 [実機単位・符号付き]; [37] IN37 B(右側) RCON1_4 SF/NG2送り 予約（使用禁止）; [38] IN38 B(右側) RCON1_4 SF/NG2送り 軸異常コード; [39] IN39 B(右側) RCON1_4 SF/NG2送り 状態信号（PEND/SV等）; [40] IN40 A(左側) RCON1_5 SF/NG2上下降 現在位置 下位 [0.01mm]; [41] IN41 A(左側) RCON1_5 SF/NG2上下降 現在位置 上位 [0.01mm]; [42] IN42 A(左側) RCON1_5 SF/NG2上下降 指令電流 下位 [mA]; [43] IN43 A(左側) RCON1_5 SF/NG2上下降 指令電流 上位 [mA]; [44] IN44 A(左側) RCON1_5 SF/NG2上下降 現在速度 [実機単位・符号付き]; [45] IN45 A(左側) RCON1_5 SF/NG2上下降 予約（使用禁止）; [46] IN46 A(左側) RCON1_5 SF/NG2上下降 軸異常コード; [47] IN47 A(左側) RCON1_5 SF/NG2上下降 状態信号（PEND/SV等）; [48] IN48 B(右側) RCON1_6 SF/NG2上下降 現在位置 下位 [0.01mm]; [49] IN49 B(右側) RCON1_6 SF/NG2上下降 現在位置 上位 [0.01mm]; [50] IN50 B(右側) RCON1_6 SF/NG2上下降 指令電流 下位 [mA]; [51] IN51 B(右側) RCON1_6 SF/NG2上下降 指令電流 上位 [mA]; [52] IN52 B(右側) RCON1_6 SF/NG2上下降 現在速度 [実機単位・符号付き]; [53] IN53 B(右側) RCON1_6 SF/NG2上下降 予約（使用禁止）; [54] IN54 B(右側) RCON1_6 SF/NG2上下降 軸異常コード; [55] IN55 B(右側) RCON1_6 SF/NG2上下降 状態信号（PEND/SV等） *)
    RCON1_TxWord : ARRAY[0..55] OF WORD;  (* 送信ワード候補; [0] OUT00 共通制御（MON/RTE）; [1] OUT01 予約（書込禁止）; [2] OUT02 予約（書込禁止）; [3] OUT03 予約（書込禁止）; [4] OUT04 予約（書込禁止）; [5] OUT05 予約（書込禁止）; [6] OUT06 予約（書込禁止）; [7] OUT07 予約（書込禁止）; [8] OUT08 A(左側) RCON1_1 NG1上下降 目標位置 下位 [0.01mm]; [9] OUT09 A(左側) RCON1_1 NG1上下降 目標位置 上位 [0.01mm]; [10] OUT10 A(左側) RCON1_1 NG1上下降 位置決め幅 下位 [0.01mm]; [11] OUT11 A(左側) RCON1_1 NG1上下降 位置決め幅 上位 [0.01mm]; [12] OUT12 A(左側) RCON1_1 NG1上下降 速度指令 [実機単位]; [13] OUT13 A(左側) RCON1_1 NG1上下降 共通加減速 [0.01G]; [14] OUT14 A(左側) RCON1_1 NG1上下降 押付け制限 [255=100%]; [15] OUT15 A(左側) RCON1_1 NG1上下降 制御信号（DSTR/SON等）; [16] OUT16 B(右側) RCON1_2 NG1上下降 目標位置 下位 [0.01mm]; [17] OUT17 B(右側) RCON1_2 NG1上下降 目標位置 上位 [0.01mm]; [18] OUT18 B(右側) RCON1_2 NG1上下降 位置決め幅 下位 [0.01mm]; [19] OUT19 B(右側) RCON1_2 NG1上下降 位置決め幅 上位 [0.01mm]; [20] OUT20 B(右側) RCON1_2 NG1上下降 速度指令 [実機単位]; [21] OUT21 B(右側) RCON1_2 NG1上下降 共通加減速 [0.01G]; [22] OUT22 B(右側) RCON1_2 NG1上下降 押付け制限 [255=100%]; [23] OUT23 B(右側) RCON1_2 NG1上下降 制御信号（DSTR/SON等）; [24] OUT24 A(左側) RCON1_3 SF/NG2仕分け(左右) 目標位置 下位 [0.01mm]; [25] OUT25 A(左側) RCON1_3 SF/NG2仕分け(左右) 目標位置 上位 [0.01mm]; [26] OUT26 A(左側) RCON1_3 SF/NG2仕分け(左右) 位置決め幅 下位 [0.01mm]; [27] OUT27 A(左側) RCON1_3 SF/NG2仕分け(左右) 位置決め幅 上位 [0.01mm]; [28] OUT28 A(左側) RCON1_3 SF/NG2仕分け(左右) 速度指令 [実機単位]; [29] OUT29 A(左側) RCON1_3 SF/NG2仕分け(左右) 共通加減速 [0.01G]; [30] OUT30 A(左側) RCON1_3 SF/NG2仕分け(左右) 押付け制限 [255=100%]; [31] OUT31 A(左側) RCON1_3 SF/NG2仕分け(左右) 制御信号（DSTR/SON等）; [32] OUT32 B(右側) RCON1_4 SF/NG2送り 目標位置 下位 [0.01mm]; [33] OUT33 B(右側) RCON1_4 SF/NG2送り 目標位置 上位 [0.01mm]; [34] OUT34 B(右側) RCON1_4 SF/NG2送り 位置決め幅 下位 [0.01mm]; [35] OUT35 B(右側) RCON1_4 SF/NG2送り 位置決め幅 上位 [0.01mm]; [36] OUT36 B(右側) RCON1_4 SF/NG2送り 速度指令 [実機単位]; [37] OUT37 B(右側) RCON1_4 SF/NG2送り 共通加減速 [0.01G]; [38] OUT38 B(右側) RCON1_4 SF/NG2送り 押付け制限 [255=100%]; [39] OUT39 B(右側) RCON1_4 SF/NG2送り 制御信号（DSTR/SON等）; [40] OUT40 A(左側) RCON1_5 SF/NG2上下降 目標位置 下位 [0.01mm]; [41] OUT41 A(左側) RCON1_5 SF/NG2上下降 目標位置 上位 [0.01mm]; [42] OUT42 A(左側) RCON1_5 SF/NG2上下降 位置決め幅 下位 [0.01mm]; [43] OUT43 A(左側) RCON1_5 SF/NG2上下降 位置決め幅 上位 [0.01mm]; [44] OUT44 A(左側) RCON1_5 SF/NG2上下降 速度指令 [実機単位]; [45] OUT45 A(左側) RCON1_5 SF/NG2上下降 共通加減速 [0.01G]; [46] OUT46 A(左側) RCON1_5 SF/NG2上下降 押付け制限 [255=100%]; [47] OUT47 A(左側) RCON1_5 SF/NG2上下降 制御信号（DSTR/SON等）; [48] OUT48 B(右側) RCON1_6 SF/NG2上下降 目標位置 下位 [0.01mm]; [49] OUT49 B(右側) RCON1_6 SF/NG2上下降 目標位置 上位 [0.01mm]; [50] OUT50 B(右側) RCON1_6 SF/NG2上下降 位置決め幅 下位 [0.01mm]; [51] OUT51 B(右側) RCON1_6 SF/NG2上下降 位置決め幅 上位 [0.01mm]; [52] OUT52 B(右側) RCON1_6 SF/NG2上下降 速度指令 [実機単位]; [53] OUT53 B(右側) RCON1_6 SF/NG2上下降 共通加減速 [0.01G]; [54] OUT54 B(右側) RCON1_6 SF/NG2上下降 押付け制限 [255=100%]; [55] OUT55 B(右側) RCON1_6 SF/NG2上下降 制御信号（DSTR/SON等） *)
    RCON1_TxUInt : ARRAY[0..55] OF UINT;  (* 送信UINT候補（実I/Oではない）; [0] OUT00 共通制御（MON/RTE）; [1] OUT01 予約（書込禁止）; [2] OUT02 予約（書込禁止）; [3] OUT03 予約（書込禁止）; [4] OUT04 予約（書込禁止）; [5] OUT05 予約（書込禁止）; [6] OUT06 予約（書込禁止）; [7] OUT07 予約（書込禁止）; [8] OUT08 A(左側) RCON1_1 NG1上下降 目標位置 下位 [0.01mm]; [9] OUT09 A(左側) RCON1_1 NG1上下降 目標位置 上位 [0.01mm]; [10] OUT10 A(左側) RCON1_1 NG1上下降 位置決め幅 下位 [0.01mm]; [11] OUT11 A(左側) RCON1_1 NG1上下降 位置決め幅 上位 [0.01mm]; [12] OUT12 A(左側) RCON1_1 NG1上下降 速度指令 [実機単位]; [13] OUT13 A(左側) RCON1_1 NG1上下降 共通加減速 [0.01G]; [14] OUT14 A(左側) RCON1_1 NG1上下降 押付け制限 [255=100%]; [15] OUT15 A(左側) RCON1_1 NG1上下降 制御信号（DSTR/SON等）; [16] OUT16 B(右側) RCON1_2 NG1上下降 目標位置 下位 [0.01mm]; [17] OUT17 B(右側) RCON1_2 NG1上下降 目標位置 上位 [0.01mm]; [18] OUT18 B(右側) RCON1_2 NG1上下降 位置決め幅 下位 [0.01mm]; [19] OUT19 B(右側) RCON1_2 NG1上下降 位置決め幅 上位 [0.01mm]; [20] OUT20 B(右側) RCON1_2 NG1上下降 速度指令 [実機単位]; [21] OUT21 B(右側) RCON1_2 NG1上下降 共通加減速 [0.01G]; [22] OUT22 B(右側) RCON1_2 NG1上下降 押付け制限 [255=100%]; [23] OUT23 B(右側) RCON1_2 NG1上下降 制御信号（DSTR/SON等）; [24] OUT24 A(左側) RCON1_3 SF/NG2仕分け(左右) 目標位置 下位 [0.01mm]; [25] OUT25 A(左側) RCON1_3 SF/NG2仕分け(左右) 目標位置 上位 [0.01mm]; [26] OUT26 A(左側) RCON1_3 SF/NG2仕分け(左右) 位置決め幅 下位 [0.01mm]; [27] OUT27 A(左側) RCON1_3 SF/NG2仕分け(左右) 位置決め幅 上位 [0.01mm]; [28] OUT28 A(左側) RCON1_3 SF/NG2仕分け(左右) 速度指令 [実機単位]; [29] OUT29 A(左側) RCON1_3 SF/NG2仕分け(左右) 共通加減速 [0.01G]; [30] OUT30 A(左側) RCON1_3 SF/NG2仕分け(左右) 押付け制限 [255=100%]; [31] OUT31 A(左側) RCON1_3 SF/NG2仕分け(左右) 制御信号（DSTR/SON等）; [32] OUT32 B(右側) RCON1_4 SF/NG2送り 目標位置 下位 [0.01mm]; [33] OUT33 B(右側) RCON1_4 SF/NG2送り 目標位置 上位 [0.01mm]; [34] OUT34 B(右側) RCON1_4 SF/NG2送り 位置決め幅 下位 [0.01mm]; [35] OUT35 B(右側) RCON1_4 SF/NG2送り 位置決め幅 上位 [0.01mm]; [36] OUT36 B(右側) RCON1_4 SF/NG2送り 速度指令 [実機単位]; [37] OUT37 B(右側) RCON1_4 SF/NG2送り 共通加減速 [0.01G]; [38] OUT38 B(右側) RCON1_4 SF/NG2送り 押付け制限 [255=100%]; [39] OUT39 B(右側) RCON1_4 SF/NG2送り 制御信号（DSTR/SON等）; [40] OUT40 A(左側) RCON1_5 SF/NG2上下降 目標位置 下位 [0.01mm]; [41] OUT41 A(左側) RCON1_5 SF/NG2上下降 目標位置 上位 [0.01mm]; [42] OUT42 A(左側) RCON1_5 SF/NG2上下降 位置決め幅 下位 [0.01mm]; [43] OUT43 A(左側) RCON1_5 SF/NG2上下降 位置決め幅 上位 [0.01mm]; [44] OUT44 A(左側) RCON1_5 SF/NG2上下降 速度指令 [実機単位]; [45] OUT45 A(左側) RCON1_5 SF/NG2上下降 共通加減速 [0.01G]; [46] OUT46 A(左側) RCON1_5 SF/NG2上下降 押付け制限 [255=100%]; [47] OUT47 A(左側) RCON1_5 SF/NG2上下降 制御信号（DSTR/SON等）; [48] OUT48 B(右側) RCON1_6 SF/NG2上下降 目標位置 下位 [0.01mm]; [49] OUT49 B(右側) RCON1_6 SF/NG2上下降 目標位置 上位 [0.01mm]; [50] OUT50 B(右側) RCON1_6 SF/NG2上下降 位置決め幅 下位 [0.01mm]; [51] OUT51 B(右側) RCON1_6 SF/NG2上下降 位置決め幅 上位 [0.01mm]; [52] OUT52 B(右側) RCON1_6 SF/NG2上下降 速度指令 [実機単位]; [53] OUT53 B(右側) RCON1_6 SF/NG2上下降 共通加減速 [0.01G]; [54] OUT54 B(右側) RCON1_6 SF/NG2上下降 押付け制限 [255=100%]; [55] OUT55 B(右側) RCON1_6 SF/NG2上下降 制御信号（DSTR/SON等） *)
    RCON1_LayoutConfirmed : BOOL;  (* I/O配置確認済み（初期OFF） *)
    RCON1_ByteOrderConfirmed : BOOL;  (* ワード・バイト順確認済み（初期OFF） *)
    RCON1_SwapBytes : BOOL;  (* 上下バイト交換設定（ON=交換） *)
    RCON1_CommOK : BOOL;  (* 通信正常（外部判定・固定ON不可） *)
    RCON1_GwMON_Request : BOOL;  (* MON要求（b15） *)
    RCON1_GwRTE_Request : BOOL;  (* 通信異常ラッチ解除要求（b13） *)
    RCON1_GwRun : BOOL;  (* GW動作中（RUN/b15） *)
    RCON1_GwControllerCommLatch : BOOL;  (* GW通信異常保持（LERC/b14） *)
    RCON1_GwAxisCommError : BOOL;  (* GW－軸 通信異常（ERRT/b13） *)
    RCON1_GwManual : BOOL;  (* 手動モード（MOD/b12） *)
    RCON1_GwHeavyAlarm : BOOL;  (* GW重故障（ALMH/b11） *)
    RCON1_GwLightAlarm : BOOL;  (* GW軽故障（ALML/b10） *)
    RCON1_GwSystemStop : BOOL;  (* システム停止状態（SEMG/b8・監視用） *)
    RCON1_GwAlarmCode : UINT;  (* GW異常コード（ALMC/b0～7） *)
    RCON1_AxisLinked : ARRAY[1..6] OF BOOL;  (* 軸別リンク状態; [1] リンク状態; [2] リンク状態; [3] リンク状態; [4] リンク状態; [5] リンク状態; [6] リンク状態 *)
    RCON1_PowerStateRaw : ARRAY[0..4] OF WORD;  (* 電源状態ワード（詳細未確認）; [0] IN02 電源状態0（詳細未確認）; [1] IN03 電源状態1（詳細未確認）; [2] IN04 電源状態2（詳細未確認）; [3] IN05 電源状態3（詳細未確認）; [4] IN06 電源状態4（詳細未確認） *)
    RCON1_EncodeOK : ARRAY[1..6] OF BOOL;  (* 軸別変換正常（運転許可とは別）; [1] 変換正常; [2] 変換正常; [3] 変換正常; [4] 変換正常; [5] 変換正常; [6] 変換正常 *)
    RCON1_EncodeError : ARRAY[1..6] OF UINT;  (* 軸別変換エラー番号（0=正常）; [1] 変換エラー番号; [2] 変換エラー番号; [3] 変換エラー番号; [4] 変換エラー番号; [5] 変換エラー番号; [6] 変換エラー番号 *)
    RCON1_WriteEnable : BOOL;  (* 実出力書込み許可（OFF=前値保持・停止不可） *)
    RCON1_GwApply : BOOL;  (* 共通出力更新許可（OFF=前値保持） *)
    RCON1_AxisApply : ARRAY[1..6] OF BOOL;  (* 軸別出力更新許可（OFF=前値保持）; [1] 出力更新許可（OFF=前値保持）; [2] 出力更新許可（OFF=前値保持）; [3] 出力更新許可（OFF=前値保持）; [4] 出力更新許可（OFF=前値保持）; [5] 出力更新許可（OFF=前値保持）; [6] 出力更新許可（OFF=前値保持） *)
    RCON1_MotionPermit : ARRAY[1..6] OF BOOL;  (* 軸別運転許可（外部判定・初期OFF）; [1] 運転許可（外部判定）; [2] 運転許可（外部判定）; [3] 運転許可（外部判定）; [4] 運転許可（外部判定）; [5] 運転許可（外部判定）; [6] 運転許可（外部判定） *)
    RCON1_GwWritten : BOOL;  (* 共通出力代入済み（RCON受付とは別） *)
    RCON1_AxisWritten : ARRAY[1..6] OF BOOL;  (* 軸別出力代入済み（RCON受付とは別）; [1] 出力代入済み（RCON受付とは別）; [2] 出力代入済み（RCON受付とは別）; [3] 出力代入済み（RCON受付とは別）; [4] 出力代入済み（RCON受付とは別）; [5] 出力代入済み（RCON受付とは別）; [6] 出力代入済み（RCON受付とは別） *)
    RCON2_RxRaw : ARRAY[0..55] OF UINT;  (* 受信値（バイト交換前）; [0] IN00 GW状態; [1] IN01 軸リンク状態; [2] IN02 電源状態0; [3] IN03 電源状態1; [4] IN04 電源状態2; [5] IN05 電源状態3; [6] IN06 電源状態4（構成依存）; [7] IN07 予約（使用禁止）; [8] IN08 1軸目 現在位置 下位 [0.01mm]; [9] IN09 1軸目 現在位置 上位 [0.01mm]; [10] IN10 1軸目 指令電流 下位 [mA]; [11] IN11 1軸目 指令電流 上位 [mA]; [12] IN12 1軸目 現在速度 [実機単位・符号付き]; [13] IN13 1軸目 予約（使用禁止）; [14] IN14 1軸目 軸異常コード; [15] IN15 1軸目 状態信号（PEND/SV等）; [16] IN16 2軸目 現在位置 下位 [0.01mm]; [17] IN17 2軸目 現在位置 上位 [0.01mm]; [18] IN18 2軸目 指令電流 下位 [mA]; [19] IN19 2軸目 指令電流 上位 [mA]; [20] IN20 2軸目 現在速度 [実機単位・符号付き]; [21] IN21 2軸目 予約（使用禁止）; [22] IN22 2軸目 軸異常コード; [23] IN23 2軸目 状態信号（PEND/SV等）; [24] IN24 3軸目 現在位置 下位 [0.01mm]; [25] IN25 3軸目 現在位置 上位 [0.01mm]; [26] IN26 3軸目 指令電流 下位 [mA]; [27] IN27 3軸目 指令電流 上位 [mA]; [28] IN28 3軸目 現在速度 [実機単位・符号付き]; [29] IN29 3軸目 予約（使用禁止）; [30] IN30 3軸目 軸異常コード; [31] IN31 3軸目 状態信号（PEND/SV等）; [32] IN32 4軸目 現在位置 下位 [0.01mm]; [33] IN33 4軸目 現在位置 上位 [0.01mm]; [34] IN34 4軸目 指令電流 下位 [mA]; [35] IN35 4軸目 指令電流 上位 [mA]; [36] IN36 4軸目 現在速度 [実機単位・符号付き]; [37] IN37 4軸目 予約（使用禁止）; [38] IN38 4軸目 軸異常コード; [39] IN39 4軸目 状態信号（PEND/SV等）; [40] IN40 5軸目 現在位置 下位 [0.01mm]; [41] IN41 5軸目 現在位置 上位 [0.01mm]; [42] IN42 5軸目 指令電流 下位 [mA]; [43] IN43 5軸目 指令電流 上位 [mA]; [44] IN44 5軸目 現在速度 [実機単位・符号付き]; [45] IN45 5軸目 予約（使用禁止）; [46] IN46 5軸目 軸異常コード; [47] IN47 5軸目 状態信号（PEND/SV等）; [48] IN48 用途未確認（今回未使用）; [49] IN49 用途未確認（今回未使用）; [50] IN50 用途未確認（今回未使用）; [51] IN51 用途未確認（今回未使用）; [52] IN52 用途未確認（今回未使用）; [53] IN53 用途未確認（今回未使用）; [54] IN54 用途未確認（今回未使用）; [55] IN55 用途未確認（今回未使用） *)
    RCON2_RxWord : ARRAY[0..55] OF WORD;  (* 受信ワード（正規化後）; [0] IN00 GW状態; [1] IN01 軸リンク状態; [2] IN02 電源状態0; [3] IN03 電源状態1; [4] IN04 電源状態2; [5] IN05 電源状態3; [6] IN06 電源状態4（構成依存）; [7] IN07 予約（使用禁止）; [8] IN08 1軸目 現在位置 下位 [0.01mm]; [9] IN09 1軸目 現在位置 上位 [0.01mm]; [10] IN10 1軸目 指令電流 下位 [mA]; [11] IN11 1軸目 指令電流 上位 [mA]; [12] IN12 1軸目 現在速度 [実機単位・符号付き]; [13] IN13 1軸目 予約（使用禁止）; [14] IN14 1軸目 軸異常コード; [15] IN15 1軸目 状態信号（PEND/SV等）; [16] IN16 2軸目 現在位置 下位 [0.01mm]; [17] IN17 2軸目 現在位置 上位 [0.01mm]; [18] IN18 2軸目 指令電流 下位 [mA]; [19] IN19 2軸目 指令電流 上位 [mA]; [20] IN20 2軸目 現在速度 [実機単位・符号付き]; [21] IN21 2軸目 予約（使用禁止）; [22] IN22 2軸目 軸異常コード; [23] IN23 2軸目 状態信号（PEND/SV等）; [24] IN24 3軸目 現在位置 下位 [0.01mm]; [25] IN25 3軸目 現在位置 上位 [0.01mm]; [26] IN26 3軸目 指令電流 下位 [mA]; [27] IN27 3軸目 指令電流 上位 [mA]; [28] IN28 3軸目 現在速度 [実機単位・符号付き]; [29] IN29 3軸目 予約（使用禁止）; [30] IN30 3軸目 軸異常コード; [31] IN31 3軸目 状態信号（PEND/SV等）; [32] IN32 4軸目 現在位置 下位 [0.01mm]; [33] IN33 4軸目 現在位置 上位 [0.01mm]; [34] IN34 4軸目 指令電流 下位 [mA]; [35] IN35 4軸目 指令電流 上位 [mA]; [36] IN36 4軸目 現在速度 [実機単位・符号付き]; [37] IN37 4軸目 予約（使用禁止）; [38] IN38 4軸目 軸異常コード; [39] IN39 4軸目 状態信号（PEND/SV等）; [40] IN40 5軸目 現在位置 下位 [0.01mm]; [41] IN41 5軸目 現在位置 上位 [0.01mm]; [42] IN42 5軸目 指令電流 下位 [mA]; [43] IN43 5軸目 指令電流 上位 [mA]; [44] IN44 5軸目 現在速度 [実機単位・符号付き]; [45] IN45 5軸目 予約（使用禁止）; [46] IN46 5軸目 軸異常コード; [47] IN47 5軸目 状態信号（PEND/SV等）; [48] IN48 用途未確認（今回未使用）; [49] IN49 用途未確認（今回未使用）; [50] IN50 用途未確認（今回未使用）; [51] IN51 用途未確認（今回未使用）; [52] IN52 用途未確認（今回未使用）; [53] IN53 用途未確認（今回未使用）; [54] IN54 用途未確認（今回未使用）; [55] IN55 用途未確認（今回未使用） *)
    RCON2_TxWord : ARRAY[0..47] OF WORD;  (* 送信ワード候補; [0] OUT00 共通制御（MON/RTE）; [1] OUT01 予約（書込禁止）; [2] OUT02 予約（書込禁止）; [3] OUT03 予約（書込禁止）; [4] OUT04 予約（書込禁止）; [5] OUT05 予約（書込禁止）; [6] OUT06 予約（書込禁止）; [7] OUT07 予約（書込禁止）; [8] OUT08 1軸目 目標位置 下位 [0.01mm]; [9] OUT09 1軸目 目標位置 上位 [0.01mm]; [10] OUT10 1軸目 位置決め幅 下位 [0.01mm]; [11] OUT11 1軸目 位置決め幅 上位 [0.01mm]; [12] OUT12 1軸目 速度指令 [実機単位]; [13] OUT13 1軸目 共通加減速 [0.01G]; [14] OUT14 1軸目 押付け制限 [255=100%]; [15] OUT15 1軸目 制御信号（DSTR/SON等）; [16] OUT16 2軸目 目標位置 下位 [0.01mm]; [17] OUT17 2軸目 目標位置 上位 [0.01mm]; [18] OUT18 2軸目 位置決め幅 下位 [0.01mm]; [19] OUT19 2軸目 位置決め幅 上位 [0.01mm]; [20] OUT20 2軸目 速度指令 [実機単位]; [21] OUT21 2軸目 共通加減速 [0.01G]; [22] OUT22 2軸目 押付け制限 [255=100%]; [23] OUT23 2軸目 制御信号（DSTR/SON等）; [24] OUT24 3軸目 目標位置 下位 [0.01mm]; [25] OUT25 3軸目 目標位置 上位 [0.01mm]; [26] OUT26 3軸目 位置決め幅 下位 [0.01mm]; [27] OUT27 3軸目 位置決め幅 上位 [0.01mm]; [28] OUT28 3軸目 速度指令 [実機単位]; [29] OUT29 3軸目 共通加減速 [0.01G]; [30] OUT30 3軸目 押付け制限 [255=100%]; [31] OUT31 3軸目 制御信号（DSTR/SON等）; [32] OUT32 4軸目 目標位置 下位 [0.01mm]; [33] OUT33 4軸目 目標位置 上位 [0.01mm]; [34] OUT34 4軸目 位置決め幅 下位 [0.01mm]; [35] OUT35 4軸目 位置決め幅 上位 [0.01mm]; [36] OUT36 4軸目 速度指令 [実機単位]; [37] OUT37 4軸目 共通加減速 [0.01G]; [38] OUT38 4軸目 押付け制限 [255=100%]; [39] OUT39 4軸目 制御信号（DSTR/SON等）; [40] OUT40 5軸目 目標位置 下位 [0.01mm]; [41] OUT41 5軸目 目標位置 上位 [0.01mm]; [42] OUT42 5軸目 位置決め幅 下位 [0.01mm]; [43] OUT43 5軸目 位置決め幅 上位 [0.01mm]; [44] OUT44 5軸目 速度指令 [実機単位]; [45] OUT45 5軸目 共通加減速 [0.01G]; [46] OUT46 5軸目 押付け制限 [255=100%]; [47] OUT47 5軸目 制御信号（DSTR/SON等） *)
    RCON2_TxUInt : ARRAY[0..47] OF UINT;  (* 送信UINT候補（実I/Oではない）; [0] OUT00 共通制御（MON/RTE）; [1] OUT01 予約（書込禁止）; [2] OUT02 予約（書込禁止）; [3] OUT03 予約（書込禁止）; [4] OUT04 予約（書込禁止）; [5] OUT05 予約（書込禁止）; [6] OUT06 予約（書込禁止）; [7] OUT07 予約（書込禁止）; [8] OUT08 1軸目 目標位置 下位 [0.01mm]; [9] OUT09 1軸目 目標位置 上位 [0.01mm]; [10] OUT10 1軸目 位置決め幅 下位 [0.01mm]; [11] OUT11 1軸目 位置決め幅 上位 [0.01mm]; [12] OUT12 1軸目 速度指令 [実機単位]; [13] OUT13 1軸目 共通加減速 [0.01G]; [14] OUT14 1軸目 押付け制限 [255=100%]; [15] OUT15 1軸目 制御信号（DSTR/SON等）; [16] OUT16 2軸目 目標位置 下位 [0.01mm]; [17] OUT17 2軸目 目標位置 上位 [0.01mm]; [18] OUT18 2軸目 位置決め幅 下位 [0.01mm]; [19] OUT19 2軸目 位置決め幅 上位 [0.01mm]; [20] OUT20 2軸目 速度指令 [実機単位]; [21] OUT21 2軸目 共通加減速 [0.01G]; [22] OUT22 2軸目 押付け制限 [255=100%]; [23] OUT23 2軸目 制御信号（DSTR/SON等）; [24] OUT24 3軸目 目標位置 下位 [0.01mm]; [25] OUT25 3軸目 目標位置 上位 [0.01mm]; [26] OUT26 3軸目 位置決め幅 下位 [0.01mm]; [27] OUT27 3軸目 位置決め幅 上位 [0.01mm]; [28] OUT28 3軸目 速度指令 [実機単位]; [29] OUT29 3軸目 共通加減速 [0.01G]; [30] OUT30 3軸目 押付け制限 [255=100%]; [31] OUT31 3軸目 制御信号（DSTR/SON等）; [32] OUT32 4軸目 目標位置 下位 [0.01mm]; [33] OUT33 4軸目 目標位置 上位 [0.01mm]; [34] OUT34 4軸目 位置決め幅 下位 [0.01mm]; [35] OUT35 4軸目 位置決め幅 上位 [0.01mm]; [36] OUT36 4軸目 速度指令 [実機単位]; [37] OUT37 4軸目 共通加減速 [0.01G]; [38] OUT38 4軸目 押付け制限 [255=100%]; [39] OUT39 4軸目 制御信号（DSTR/SON等）; [40] OUT40 5軸目 目標位置 下位 [0.01mm]; [41] OUT41 5軸目 目標位置 上位 [0.01mm]; [42] OUT42 5軸目 位置決め幅 下位 [0.01mm]; [43] OUT43 5軸目 位置決め幅 上位 [0.01mm]; [44] OUT44 5軸目 速度指令 [実機単位]; [45] OUT45 5軸目 共通加減速 [0.01G]; [46] OUT46 5軸目 押付け制限 [255=100%]; [47] OUT47 5軸目 制御信号（DSTR/SON等） *)
    RCON2_LayoutConfirmed : BOOL;  (* I/O配置確認済み（初期OFF） *)
    RCON2_ByteOrderConfirmed : BOOL;  (* ワード・バイト順確認済み（初期OFF） *)
    RCON2_SwapBytes : BOOL;  (* 上下バイト交換設定（ON=交換） *)
    RCON2_CommOK : BOOL;  (* 通信正常（外部判定・固定ON不可） *)
    RCON2_GwMON_Request : BOOL;  (* MON要求（b15） *)
    RCON2_GwRTE_Request : BOOL;  (* 通信異常ラッチ解除要求（b13） *)
    RCON2_GwRun : BOOL;  (* GW動作中（RUN/b15） *)
    RCON2_GwControllerCommLatch : BOOL;  (* GW通信異常保持（LERC/b14） *)
    RCON2_GwAxisCommError : BOOL;  (* GW－軸 通信異常（ERRT/b13） *)
    RCON2_GwManual : BOOL;  (* 手動モード（MOD/b12） *)
    RCON2_GwHeavyAlarm : BOOL;  (* GW重故障（ALMH/b11） *)
    RCON2_GwLightAlarm : BOOL;  (* GW軽故障（ALML/b10） *)
    RCON2_GwSystemStop : BOOL;  (* システム停止状態（SEMG/b8・監視用） *)
    RCON2_GwAlarmCode : UINT;  (* GW異常コード（ALMC/b0～7） *)
    RCON2_AxisLinked : ARRAY[1..5] OF BOOL;  (* 軸別リンク状態; [1] 1軸目（No.0）リンク状態; [2] 2軸目（No.1）リンク状態; [3] 3軸目（No.2）リンク状態; [4] 4軸目（No.3）リンク状態; [5] 5軸目（No.4）リンク状態 *)
    RCON2_PowerStateRaw : ARRAY[0..4] OF WORD;  (* 電源状態ワード（詳細未確認）; [0] IN02 電源状態0（詳細未確認）; [1] IN03 電源状態1（詳細未確認）; [2] IN04 電源状態2（詳細未確認）; [3] IN05 電源状態3（詳細未確認）; [4] IN06 電源状態4（詳細未確認） *)
    RCON2_EncodeOK : ARRAY[1..5] OF BOOL;  (* 軸別変換正常（運転許可とは別）; [1] 1軸目（No.0）変換正常; [2] 2軸目（No.1）変換正常; [3] 3軸目（No.2）変換正常; [4] 4軸目（No.3）変換正常; [5] 5軸目（No.4）変換正常 *)
    RCON2_EncodeError : ARRAY[1..5] OF UINT;  (* 軸別変換エラー番号（0=正常）; [1] 1軸目（No.0）変換エラー番号; [2] 2軸目（No.1）変換エラー番号; [3] 3軸目（No.2）変換エラー番号; [4] 4軸目（No.3）変換エラー番号; [5] 5軸目（No.4）変換エラー番号 *)
    RCON2_WriteEnable : BOOL;  (* 実出力書込み許可（OFF=前値保持・停止不可） *)
    RCON2_GwApply : BOOL;  (* 共通出力更新許可（OFF=前値保持） *)
    RCON2_AxisApply : ARRAY[1..5] OF BOOL;  (* 軸別出力更新許可（OFF=前値保持）; [1] 1軸目（No.0）出力更新許可（OFF=前値保持）; [2] 2軸目（No.1）出力更新許可（OFF=前値保持）; [3] 3軸目（No.2）出力更新許可（OFF=前値保持）; [4] 4軸目（No.3）出力更新許可（OFF=前値保持）; [5] 5軸目（No.4）出力更新許可（OFF=前値保持） *)
    RCON2_MotionPermit : ARRAY[1..5] OF BOOL;  (* 軸別運転許可（外部判定・初期OFF）; [1] 1軸目（No.0）運転許可（外部判定）; [2] 2軸目（No.1）運転許可（外部判定）; [3] 3軸目（No.2）運転許可（外部判定）; [4] 4軸目（No.3）運転許可（外部判定）; [5] 5軸目（No.4）運転許可（外部判定） *)
    RCON2_GwWritten : BOOL;  (* 共通出力代入済み（RCON受付とは別） *)
    RCON2_AxisWritten : ARRAY[1..5] OF BOOL;  (* 軸別出力代入済み（RCON受付とは別）; [1] 1軸目（No.0）出力代入済み（RCON受付とは別）; [2] 2軸目（No.1）出力代入済み（RCON受付とは別）; [3] 3軸目（No.2）出力代入済み（RCON受付とは別）; [4] 4軸目（No.3）出力代入済み（RCON受付とは別）; [5] 5軸目（No.4）出力代入済み（RCON受付とは別） *)
    RCON1_1_Auto : ARRAY[0..99] OF Bool;  (* 自動移動要求; [1] 原点位置移動; [2] NG仕分け; [3] 動作完了後 原点位置移動 *)
    RCON1_1_OUT_PositionBand_mm : LREAL;  (* 位置決め幅 [mm] *)
    RCON1_1_OUT_TargetPos_mm : LREAL;  (* 目標位置 [mm] *)
    RCON1_1_OUT_Speed_mm_s : LREAL;  (* 指令速度 [mm/s] *)
    RCON1_1_OUT_AccDec_G : LREAL;  (* 加減速度 [G] *)
    RCON1_1_OUT_PushLimit_pct : LREAL;  (* 押付け制限 [%]（未使用） *)
    RCON1_1_ActualPos_mm : LREAL;  (* 現在位置 [mm] *)
    RCON1_1_Current_mA : DINT;  (* 指令電流 [mA]（監視値） *)
    RCON1_1_ActualSpeed_mm_s : LREAL;  (* 現在速度 [mm/s] *)
    RCON1_1_AlarmCode : UINT;  (* 軸異常コード *)
    RCON1_1_DataValid : BOOL;  (* 入力有効（安全許可とは別） *)
    RCON1_1_IN_PositionDone : BOOL;  (* 位置決め完了 *)
    RCON1_1_IN_HomeDone : BOOL;  (* 原点復帰完了 *)
    RCON1_1_IN_Moving : BOOL;  (* 移動中 *)
    RCON1_1_IN_EmergencyStop : BOOL;  (* 非常停止状態（監視） *)
    RCON1_1_IN_ControllerReady : BOOL;  (* 準備完了 *)
    RCON1_1_IN_Zone2 : BOOL;  (* ゾーン2内 *)
    RCON1_1_IN_Zone1 : BOOL;  (* ゾーン1内 *)
    RCON1_1_IN_CommandDone : BOOL;  (* 指令完了 *)
    RCON1_1_IN_OverloadWarning : BOOL;  (* 過負荷警告 *)
    RCON1_1_IN_PushMiss : BOOL;  (* 押付け空振り（未使用） *)
    RCON1_1_IN_ServoReady : BOOL;  (* サーボON状態 *)
    RCON1_1_IN_Alarm : BOOL;  (* 軸異常 *)
    RCON1_1_Ready : BOOL;  (* 動作準備（安全許可とは別） *)
    RCON1_1_Error : BOOL;  (* 異常予備（未接続） *)
    RCON1_1_Error_Clear : BOOL;  (* 解除予備（未接続） *)
    Error_M : ARRAY[0..99] OF Bool;  (* エラー：; [1] シリンダ; [2] コンベア＆ドアセンサ; [3] FH A(左側) ST1; [4] A(左側)検査コンベア ワーク不一致; [5] RCON1-1 異常; [6] GT2 エラー; [7] NG1仕分けエラー; [8] 反転1エラー; [9] FH A(左側) ST5; [10] FH B(右側) ST1; [11] FH B(右側) ST5; [12] A(左側) ST6 反転2 ワーク不一致; [13] ST7 排出前ワーク不一致エラー *)
    HMI_RCON1_1_OUT_TargetPos : ARRAY[0..99] OF LREAL;  (* HMI設定位置 [mm]; [1] 原点位置; [3] 高さNG位置; [4] カメラ キズNG位置; [5] カメラ 姿NG位置 *)
    RCON1_1_M : ARRAY[0..99] OF BOOL;  (* #A(左側) RCON1_1 NG1排出(上下); [1] 開始指令保持; [2] 予備 *)
    RCON1_1_MoveDone : BOOL;  (* 動作完了 *)
    ST1_A_Ca1_M : ARRAY[0..99] OF Bool;  (* [1] ST1 A カメラ1 検査開始; [2] 【Y720】A(左側) 位置1ストッパー 戻; [3] ワーク有無 判定; [4] ST1 A ワーク有; [5] ST1 A ワーク無; [6] A(左側) ST1 検査前ワーク不一致; [7] ST1 FH測定開始 *)
    ST2_A_Hgt_M : ARRAY[0..99] OF Bool;  (* [4] 【Y721】A(左側) 位置2ストッパー戻; [6] ST2 A ワーク有＆工程OK; [7] ST2 A ワーク無 or 前工程NG; [5] ワーク有無 判定; [9] 【Y703】A(左側) 高さ検査持上行; [10] 【Y701】A(左側) 高さ検査押え行; [11] A(左側) 高さ検査OK判定; [12] A(左側) 高さ検査NG判定; [2] 【Y701】A(左側) 高さ検査押え行; [8] ST2 検査前ワーク不一致エラー *)
    ST3_A_Dis1_End : BOOL;  (* ST3 A 動作完了 *)
    ST3_A_Dis1_M : ARRAY[0..99] OF Bool;  (* [7] 原点位置 移動開始; [6] 原点位置移動 データ転送; [5] 【Y722】A(左側) 位置3ストッパー戻; [4] 【Y706】A(左側) NG1チャック戻; [8] ワーク有無 / 検査前ワーク不一致 判定; [9] ST3 A ワーク有＆工程NG; [10] ST3 A ワーク無 or 前工程OK; [14] 【Y704】A(左側) NG1ピックアップ戻 ; [24] 仕分け完了; [16] 高さNG位置; [17] カメラ キズNG位置; [18] カメラ 姿NG位置; [21] 高さNG; [22] カメラ キズNG; [23] カメラ 姿NG; [11] ST3 検査前ワーク不一致エラー; [25] #動作完了後 原点位置移動; [12] 【Y705】A(左側) NG1ピックアップ 行 *)
    Homing_Para_Stm : _sHOMING_REF;
    Stm_A_Rev_Axis000_OriginDone : BOOL;  (* A(左側) ST4 反転1 モータ原点復帰完了 *)
    HMI_Home_SW : BOOL;  (* HMI 原点復帰SW *)
    Origin_Busy : BOOL;  (* 原点復帰中 *)
    Out_CYw_Rev_01_Pick_A_H_Origin : ARRAY[0..10] OF Bool;  (* 原点復帰【Y710】A(左側)ST4 反転1ピックアップ戻： *)
    Stm_A_Rev_Axis000_Origin : BOOL;  (* A(左側) ST4 反転1 モータ原点復帰開始 *)
    Out_CYw_Rev_01_Pick_A_F_Origin : ARRAY[0..99] OF Bool;  (* 原点復帰【Y711】A(左側)ST4 反転1ピックアップ行： *)
    Out_CYw_Rev_01_Chk_A_H_Origin : ARRAY[0..99] OF Bool;  (* 原点復帰【Y708】A(左側)ST4 反転1チャック閉： *)
    Stm_A_Rev_Axis001_Origin : BOOL;  (* A(左側) ST6 反転2 モータ原点復帰開始 *)
    Stm_A_Rev_Axis001_OriginDone : BOOL;  (* A(左側) ST6 反転2 モータ原点復帰完了 *)
    Out_CYw_Rev_02_Pick_A_H_Origin : ARRAY[0..10] OF Bool;  (* 原点復帰 【Y714】A(左側)ST6 反転2ピックアップ戻 *)
    Out_CYw_Rev_02_Pick_A_F_Origin : ARRAY[0..99] OF Bool;  (* 原点復帰 【Y715】A(左側)ST6 反転2ピックアップ行 *)
    Out_CYw_Rev_02_Chk_A_H_Origin : ARRAY[0..99] OF Bool;  (* 原点復帰 【Y712】A(左側)ST6 反転2チャック閉 戻 *)
    Auto_B_Start : BOOL;  (* B(右側)自動運転開始（後続処理未接続） *)
    Stm_B_Rev_Axis002_Origin : BOOL;  (* B(右側) ST4 反転1 モータ原点復帰開始 *)
    Stm_B_Rev_Axis002_OriginDone : BOOL;  (* B(右側) ST4 反転1 モータ原点復帰完了 *)
    Out_CYw_Rev_01_Pick_B_H_Origin : ARRAY[0..10] OF Bool;  (* 原点復帰 【Y810】B(右側)ST4 反転1ピックアップ戻 *)
    Out_CYw_Rev_01_Pick_B_F_Origin : ARRAY[0..99] OF Bool;  (* 原点復帰 【Y811】B(右側)ST4 反転1ピックアップ行 *)
    Out_CYw_Rev_01_Chk_B_H_Origin : ARRAY[0..99] OF Bool;  (* 原点復帰 【Y808】B(右側)ST4 反転1チャック閉 戻 *)
    Stm_B_Rev_Axis003_Origin : BOOL;  (* B(右側) ST6 反転2 モータ原点復帰開始 *)
    Stm_B_Rev_Axis003_OriginDone : BOOL;  (* B(右側) ST6 反転2 モータ原点復帰完了 *)
    Out_CYw_Rev_02_Pick_B_H_Origin : ARRAY[0..10] OF Bool;  (* 原点復帰 【Y814】B(右側)ST6 反転2ピックアップ戻 *)
    Out_CYw_Rev_02_Pick_B_F_Origin : ARRAY[0..99] OF Bool;  (* 原点復帰 【Y815】B(右側)ST6 反転2ピックアップ行 *)
    Out_CYw_Rev_02_Chk_B_H_Origin : ARRAY[0..99] OF Bool;  (* 原点復帰 【Y812】B(右側)ST6 反転2チャック閉 戻 *)
    E001_Out_OUT00_2003_01_1 : UINT;
    ST4_A_Rev1_M : ARRAY[0..99] OF Bool;  (* [2] 【Y710】A(左側)ST4 反転1ピックアップ戻; [3] 【Y723】A(左側) 位置4ストッパー戻; [4] 原点位置移動 データ転送; [5] 原点位置移動 開始; [6] A(左側)ステッピング反転モータ1 絶対値位置決め 動作完了; [7] ワーク有無 / 検査前ワーク不一致 判定; [8] ST4 A ワーク有＆工程OK; [9] ST4 A ワーク無 or 前工程NG; [10] A(左側) ST4 ワーク不一致エラー; [12] 【Y708】A(左側) ST4 反転1チャック閉; [13] 【Y710】A(左側)ST4 反転1ピックアップ戻; [14] 原点位置移動(180°) データ転送; [15] A(左側)ステッピング反転モータ1 絶対値位置決め 動作完了; [16] 【Y711】A(左側)ST4 反転1ピックアップ行; [17] 【Y709】A(左側)ST4 反転1チャック開 行; [18] 【Y710】A(左側)ST4 反転1ピックアップ戻 *)
    Stm_A_Rev_Axis000_MovePos_Degree : LREAL;  (* A(左側)ステッピングモータ000 回転角度 *)
    Stm_A_Rev_Axis000_MoveAbsoluteDone : BOOL;  (* A(左側)ステッピング反転モータ1 絶対値位置決め 動作完了 *)
    HMI_Stm_A_Rev_Axis000_MovePos_Degree : ARRAY[0..99] OF LREAL;  (* A(左側)ステッピングモータ000 回転角度; [2] ワーク反転動作 *)
    Stm_A_Rev_Axis000_Auto : ARRAY[0..99] OF Bool;  (* [1] 原点位置移動 開始 *)
    ST5_A_Ca2_M : ARRAY[0..99] OF Bool;  (* [1] A(左側) ST5 カメラ2検査開始; [2] 【Y724】A(左側) ST5 ストッパー戻; [3] A(左側) ST5 ワーク有無判定; [4] A(左側) ST5 ワーク有; [5] A(左側) ST5 ワーク無; [6] A(左側) ST5 検査前ワーク不一致; [7] A(左側) ST5 FH測定開始 *)
    ST5_A_Ca2_Busy : BOOL;  (* A(左側) ST5 カメラ2検査中 *)
    ST5_A_Ca2_End : BOOL;  (* A(左側) ST5 カメラ2動作完了 *)
    FH_A_ST5_Auto : BOOL;  (* A(左側) ST5 FH自動測定 *)
    FH_A_ST5_Manual : BOOL;  (* A(左側) ST5 FH手動測定 *)
    FH_A_ST5_Done : BOOL;  (* A(左側) ST5 画像検査完了 *)
    ST6_A_Rev2_M : ARRAY[0..99] OF Bool;  (* [1] A(左側) ST6 反転2 動作開始; [2] A(左側) ST6 反転2 【Y714】ピックアップ戻; [3] A(左側) ST6 反転2 【Y725】位置6ストッパー戻; [4] A(左側) ST6 反転2 原点角度転送; [5] A(左側) ST6 反転2 原点位置移動開始; [6] A(左側) ST6 反転2 原点位置移動完了; [7] A(左側) ST6 反転2 ワーク有無判定; [8] A(左側) ST6 反転2 ワーク有・前工程OK; [9] A(左側) ST6 反転2 ワーク無・前工程NG; [10] A(左側) ST6 反転2 ワーク不一致; [11] A(左側) ST6 反転2 【Y715】反転前ピックアップ行; [12] A(左側) ST6 反転2 【Y712】チャック閉; [13] A(左側) ST6 反転2 【Y714】反転前ピックアップ戻; [14] A(左側) ST6 反転2 反転角度転送; [15] A(左側) ST6 反転2 反転位置移動完了; [16] A(左側) ST6 反転2 【Y715】設置ピックアップ行; [17] A(左側) ST6 反転2 【Y713】チャック開; [18] A(左側) ST6 反転2 【Y714】設置ピックアップ戻 *)
    Stm_A_Rev_Axis001_MovePos_Degree : LREAL;  (* A(左側) ST6 反転2指令角度 *)
    Stm_A_Rev_Axis001_MoveAbsoluteDone : BOOL;  (* A(左側) ST6 反転2位置決め完了 *)
    HMI_Stm_A_Rev_Axis001_MovePos_Degree : ARRAY[0..99] OF LREAL;  (* A(左側) ST6 反転2設定角度; [1] A(左側) ST6 原点位置設定角度; [2] A(左側) ST6 反転位置設定角度 *)
    Stm_A_Rev_Axis001_Auto : ARRAY[0..99] OF Bool;  (* A(左側) ST6 反転2自動指令; [1] A(左側) ST6 原点位置移動開始 *)
    Homing_Para_Stm_Rev2 : _sHOMING_REF;  (* A(左側) ST6 反転2原点設定 *)
    RCON1_2_IN_PositionDone : BOOL;  (* 位置決め完了 *)
    RCON1_2_IN_HomeDone : BOOL;  (* 原点復帰完了 *)
    RCON1_2_IN_Moving : BOOL;  (* 移動中 *)
    RCON1_2_IN_EmergencyStop : BOOL;  (* 非常停止状態（監視） *)
    RCON1_2_IN_ControllerReady : BOOL;  (* 準備完了 *)
    RCON1_2_IN_Zone2 : BOOL;  (* ゾーン2内 *)
    RCON1_2_IN_Zone1 : BOOL;  (* ゾーン1内 *)
    RCON1_2_IN_CommandDone : BOOL;  (* 指令完了 *)
    RCON1_2_IN_OverloadWarning : BOOL;  (* 過負荷警告 *)
    RCON1_2_IN_PushMiss : BOOL;  (* 押付け空振り（未使用） *)
    RCON1_2_IN_ServoReady : BOOL;  (* サーボON状態 *)
    RCON1_2_IN_Alarm : BOOL;  (* 軸異常 *)
    RCON1_2_Ready : BOOL;  (* 動作準備（安全許可とは別） *)
    RCON1_2_Error : BOOL;  (* 異常予備（未接続） *)
    RCON1_2_Error_Clear : BOOL;  (* 解除予備（未接続） *)
    RCON1_2_M : ARRAY[0..99] OF BOOL;  (* #B(右側) RCON1_2 NG1排出(上下); [1] 開始指令保持; [2] 予備 *)
    RCON1_2_MoveDone : BOOL;  (* 動作完了 *)
    RCON1_2_OUT_TargetPos_mm : LREAL;  (* 目標位置 [mm] *)
    RCON1_2_OUT_PositionBand_mm : LREAL;  (* 位置決め幅 [mm] *)
    RCON1_2_OUT_Speed_mm_s : LREAL;  (* 指令速度 [mm/s] *)
    RCON1_2_OUT_AccDec_G : LREAL;  (* 加減速度 [G] *)
    RCON1_2_OUT_PushLimit_pct : LREAL;  (* 押付け制限 [%]（未使用） *)
    RCON1_2_ActualPos_mm : LREAL;  (* 現在位置 [mm] *)
    RCON1_2_Current_mA : DINT;  (* 指令電流 [mA]（監視値） *)
    RCON1_2_ActualSpeed_mm_s : LREAL;  (* 現在速度 [mm/s] *)
    RCON1_2_AlarmCode : UINT;  (* 軸異常コード *)
    RCON1_2_DataValid : BOOL;  (* 入力有効（安全許可とは別） *)
    RCON1_2_Auto : ARRAY[0..99] OF Bool;  (* 自動移動要求; [1] 自動要求1（外部接続用）; [2] 自動要求2（外部接続用）; [3] 自動要求3（外部接続用） *)
    RCON1_3_IN_PositionDone : BOOL;  (* 位置決め完了 *)
    RCON1_3_IN_HomeDone : BOOL;  (* 原点復帰完了 *)
    RCON1_3_IN_Moving : BOOL;  (* 移動中 *)
    RCON1_3_IN_EmergencyStop : BOOL;  (* 非常停止状態（監視） *)
    RCON1_3_IN_ControllerReady : BOOL;  (* 準備完了 *)
    RCON1_3_IN_Zone2 : BOOL;  (* ゾーン2内 *)
    RCON1_3_IN_Zone1 : BOOL;  (* ゾーン1内 *)
    RCON1_3_IN_CommandDone : BOOL;  (* 指令完了 *)
    RCON1_3_IN_OverloadWarning : BOOL;  (* 過負荷警告 *)
    RCON1_3_IN_PushMiss : BOOL;  (* 押付け空振り（未使用） *)
    RCON1_3_IN_ServoReady : BOOL;  (* サーボON状態 *)
    RCON1_3_IN_Alarm : BOOL;  (* 軸異常 *)
    RCON1_3_Ready : BOOL;  (* 動作準備（安全許可とは別） *)
    RCON1_3_Error : BOOL;  (* 異常予備（未接続） *)
    RCON1_3_Error_Clear : BOOL;  (* 解除予備（未接続） *)
    RCON1_3_M : ARRAY[0..99] OF BOOL;  (* #A(左側) RCON1_3 SF/NG2仕分け(左右); [1] 開始指令保持; [2] 予備 *)
    RCON1_3_MoveDone : BOOL;  (* 動作完了 *)
    RCON1_3_OUT_TargetPos_mm : LREAL;  (* 目標位置 [mm] *)
    RCON1_3_OUT_PositionBand_mm : LREAL;  (* 位置決め幅 [mm] *)
    RCON1_3_OUT_Speed_mm_s : LREAL;  (* 指令速度 [mm/s] *)
    RCON1_3_OUT_AccDec_G : LREAL;  (* 加減速度 [G] *)
    RCON1_3_OUT_PushLimit_pct : LREAL;  (* 押付け制限 [%]（未使用） *)
    RCON1_3_ActualPos_mm : LREAL;  (* 現在位置 [mm] *)
    RCON1_3_Current_mA : DINT;  (* 指令電流 [mA]（監視値） *)
    RCON1_3_ActualSpeed_mm_s : LREAL;  (* 現在速度 [mm/s] *)
    RCON1_3_AlarmCode : UINT;  (* 軸異常コード *)
    RCON1_3_DataValid : BOOL;  (* 入力有効（安全許可とは別） *)
    RCON1_3_Auto : ARRAY[0..99] OF Bool;  (* 自動移動要求; [1] 原点位置移動; [2] 自動要求2（外部接続用）; [3] 自動要求3（外部接続用） *)
    RCON1_4_IN_PositionDone : BOOL;  (* 位置決め完了 *)
    RCON1_4_IN_HomeDone : BOOL;  (* 原点復帰完了 *)
    RCON1_4_IN_Moving : BOOL;  (* 移動中 *)
    RCON1_4_IN_EmergencyStop : BOOL;  (* 非常停止状態（監視） *)
    RCON1_4_IN_ControllerReady : BOOL;  (* 準備完了 *)
    RCON1_4_IN_Zone2 : BOOL;  (* ゾーン2内 *)
    RCON1_4_IN_Zone1 : BOOL;  (* ゾーン1内 *)
    RCON1_4_IN_CommandDone : BOOL;  (* 指令完了 *)
    RCON1_4_IN_OverloadWarning : BOOL;  (* 過負荷警告 *)
    RCON1_4_IN_PushMiss : BOOL;  (* 押付け空振り（未使用） *)
    RCON1_4_IN_ServoReady : BOOL;  (* サーボON状態 *)
    RCON1_4_IN_Alarm : BOOL;  (* 軸異常 *)
    RCON1_4_Ready : BOOL;  (* 動作準備（安全許可とは別） *)
    RCON1_4_Error : BOOL;  (* 異常予備（未接続） *)
    RCON1_4_Error_Clear : BOOL;  (* 解除予備（未接続） *)
    RCON1_4_M : ARRAY[0..99] OF BOOL;  (* #B(右側) RCON1_4 SF/NG2排出(送り); [1] 開始指令保持; [2] 予備 *)
    RCON1_4_MoveDone : BOOL;  (* 動作完了 *)
    RCON1_4_OUT_TargetPos_mm : LREAL;  (* 目標位置 [mm] *)
    RCON1_4_OUT_PositionBand_mm : LREAL;  (* 位置決め幅 [mm] *)
    RCON1_4_OUT_Speed_mm_s : LREAL;  (* 指令速度 [mm/s] *)
    RCON1_4_OUT_AccDec_G : LREAL;  (* 加減速度 [G] *)
    RCON1_4_OUT_PushLimit_pct : LREAL;  (* 押付け制限 [%]（未使用） *)
    RCON1_4_ActualPos_mm : LREAL;  (* 現在位置 [mm] *)
    RCON1_4_Current_mA : DINT;  (* 指令電流 [mA]（監視値） *)
    RCON1_4_ActualSpeed_mm_s : LREAL;  (* 現在速度 [mm/s] *)
    RCON1_4_AlarmCode : UINT;  (* 軸異常コード *)
    RCON1_4_DataValid : BOOL;  (* 入力有効（安全許可とは別） *)
    RCON1_4_Auto : ARRAY[0..99] OF Bool;  (* 自動移動要求; [1] 自動要求1（外部接続用）; [2] 自動要求2（外部接続用）; [3] 自動要求3（外部接続用） *)
    RCON1_5_IN_PositionDone : BOOL;  (* 位置決め完了 *)
    RCON1_5_IN_HomeDone : BOOL;  (* 原点復帰完了 *)
    RCON1_5_IN_Moving : BOOL;  (* 移動中 *)
    RCON1_5_IN_EmergencyStop : BOOL;  (* 非常停止状態（監視） *)
    RCON1_5_IN_ControllerReady : BOOL;  (* 準備完了 *)
    RCON1_5_IN_Zone2 : BOOL;  (* ゾーン2内 *)
    RCON1_5_IN_Zone1 : BOOL;  (* ゾーン1内 *)
    RCON1_5_IN_CommandDone : BOOL;  (* 指令完了 *)
    RCON1_5_IN_OverloadWarning : BOOL;  (* 過負荷警告 *)
    RCON1_5_IN_PushMiss : BOOL;  (* 押付け空振り（未使用） *)
    RCON1_5_IN_ServoReady : BOOL;  (* サーボON状態 *)
    RCON1_5_IN_Alarm : BOOL;  (* 軸異常 *)
    RCON1_5_Ready : BOOL;  (* 動作準備（安全許可とは別） *)
    RCON1_5_Error : BOOL;  (* 異常予備（未接続） *)
    RCON1_5_Error_Clear : BOOL;  (* 解除予備（未接続） *)
    RCON1_5_M : ARRAY[0..99] OF BOOL;  (* #A(左側) RCON1_5 SF/NG2排出(上下); [1] 開始指令保持; [2] 予備 *)
    RCON1_5_MoveDone : BOOL;  (* 動作完了 *)
    RCON1_5_OUT_TargetPos_mm : LREAL;  (* 目標位置 [mm] *)
    RCON1_5_OUT_PositionBand_mm : LREAL;  (* 位置決め幅 [mm] *)
    RCON1_5_OUT_Speed_mm_s : LREAL;  (* 指令速度 [mm/s] *)
    RCON1_5_OUT_AccDec_G : LREAL;  (* 加減速度 [G] *)
    RCON1_5_OUT_PushLimit_pct : LREAL;  (* 押付け制限 [%]（未使用） *)
    RCON1_5_ActualPos_mm : LREAL;  (* 現在位置 [mm] *)
    RCON1_5_Current_mA : DINT;  (* 指令電流 [mA]（監視値） *)
    RCON1_5_ActualSpeed_mm_s : LREAL;  (* 現在速度 [mm/s] *)
    RCON1_5_AlarmCode : UINT;  (* 軸異常コード *)
    RCON1_5_DataValid : BOOL;  (* 入力有効（安全許可とは別） *)
    RCON1_5_Auto : ARRAY[0..99] OF Bool;  (* 自動移動要求; [1] 原点位置移動; [2] 自動要求2（外部接続用）; [3] 自動要求3（外部接続用） *)
    RCON1_6_IN_PositionDone : BOOL;  (* 位置決め完了 *)
    RCON1_6_IN_HomeDone : BOOL;  (* 原点復帰完了 *)
    RCON1_6_IN_Moving : BOOL;  (* 移動中 *)
    RCON1_6_IN_EmergencyStop : BOOL;  (* 非常停止状態（監視） *)
    RCON1_6_IN_ControllerReady : BOOL;  (* 準備完了 *)
    RCON1_6_IN_Zone2 : BOOL;  (* ゾーン2内 *)
    RCON1_6_IN_Zone1 : BOOL;  (* ゾーン1内 *)
    RCON1_6_IN_CommandDone : BOOL;  (* 指令完了 *)
    RCON1_6_IN_OverloadWarning : BOOL;  (* 過負荷警告 *)
    RCON1_6_IN_PushMiss : BOOL;  (* 押付け空振り（未使用） *)
    RCON1_6_IN_ServoReady : BOOL;  (* サーボON状態 *)
    RCON1_6_IN_Alarm : BOOL;  (* 軸異常 *)
    RCON1_6_Ready : BOOL;  (* 動作準備（安全許可とは別） *)
    RCON1_6_Error : BOOL;  (* 異常予備（未接続） *)
    RCON1_6_Error_Clear : BOOL;  (* 解除予備（未接続） *)
    RCON1_6_M : ARRAY[0..99] OF BOOL;  (* #B(右側) RCON1_6 SF/NG2排出(上下); [1] 開始指令保持; [2] 予備 *)
    RCON1_6_MoveDone : BOOL;  (* 動作完了 *)
    RCON1_6_OUT_TargetPos_mm : LREAL;  (* 目標位置 [mm] *)
    RCON1_6_OUT_PositionBand_mm : LREAL;  (* 位置決め幅 [mm] *)
    RCON1_6_OUT_Speed_mm_s : LREAL;  (* 指令速度 [mm/s] *)
    RCON1_6_OUT_AccDec_G : LREAL;  (* 加減速度 [G] *)
    RCON1_6_OUT_PushLimit_pct : LREAL;  (* 押付け制限 [%]（未使用） *)
    RCON1_6_ActualPos_mm : LREAL;  (* 現在位置 [mm] *)
    RCON1_6_Current_mA : DINT;  (* 指令電流 [mA]（監視値） *)
    RCON1_6_ActualSpeed_mm_s : LREAL;  (* 現在速度 [mm/s] *)
    RCON1_6_AlarmCode : UINT;  (* 軸異常コード *)
    RCON1_6_DataValid : BOOL;  (* 入力有効（安全許可とは別） *)
    RCON1_6_Auto : ARRAY[0..99] OF Bool;  (* 自動移動要求; [1] 自動要求1（外部接続用）; [2] 自動要求2（外部接続用）; [3] 自動要求3（外部接続用） *)
END_VAR
VAR_GLOBAL RETAIN
    HMI_RCON1_5_OUT_TargetPos : ARRAY[0..99] OF LREAL;  (* RCON1_5 SF/NG2排出(上下) 目標位置 [mm]：; [1] 原点位置移動 *)
    HMI_RCON1_3_OUT_TargetPos : ARRAY[0..99] OF LREAL;  (* RCON1_3 SF/NG2仕分け(左右) 目標位置 [mm]： *)
END_VAR
VAR_GLOBAL
    ST7_A_Dis2_M : ARRAY[0..99] OF Bool;  (* [9] ST7 A ワーク有; [10] ST3 A ワーク無; [11] ST7 排出前ワーク不一致エラー *)
END_VAR

